 (*Air Pressure*)
'101x003x011',   'Warning',      'Zone 1 CIP - Air pressure is Low',
'101x003x012',   'Warning',      'Zone 2 TriBlender - Air pressure is Low',
'101x003x013',   'Warning',      'Zone 3 Marinade - Air pressure is Low',
'101x003x014',   'Warning',      'Zone 4 Color - Air pressure is Low',

'101x003x021',   'Warning',      'Zone 1 CIP - Air pressure is High',
'101x003x022',   'Warning',      'Zone 2 TriBlender - Air pressure is High',
'101x003x023',   'Warning',      'Zone 3 Marinade - Air pressure is High',
'101x003x024',   'Warning',      'Zone 4 Color - Air pressure is High',

'101x003x111',   'Error',      'Zone 1 CIP - Air pressure is Low',
'101x003x112',   'Error',      'Zone 2 TriBlender - Air pressure is Low',
'101x003x113',   'Error',      'Zone 3 Marinade - Air pressure is Low',
'101x003x114',   'Error',      'Zone 4 Color - Air pressure is Low',

'101x003x121',   'Error',      'Zone 1 CIP - Air pressure is High',
'101x003x122',   'Error',      'Zone 2 TriBlender - Air pressure is High',
'101x003x123',   'Error',      'Zone 3 Marinade - Air pressure is High',
'101x003x124',   'Error',      'Zone 4 Color - Air pressure is High',


  
    (*Emergency*)
'106x001x001',   'Error',      'Emergency cycle 1 (CIP) circuit interrupted',
'106x002x001',   'Error',      'Emergency cycle 2 (Color) circuit interrupted',
'106x003x001',   'Error',      'Emergency cycle 3 (TriBlender) circuit interrupted',
'106x004x001',   'Error',      'Emergency cycle 4 (Marinade) circuit interrupted',

'106x001x002',   'Warning',    'Emergency PB1 Pressed',
'106x002x002',   'Warning',    'Emergency PB2 Pressed',
'106x003x002',   'Warning',    'Emergency PB3_1 Pressed',
'106x003x003',   'Warning',    'Emergency PB3_2 Pressed',
'106x004x002',   'Warning',    'Emergency PB4 Pressed',
'106x000x060',   'Message',    'Emergency Bypass activated',	








    (*Doors*)
	
'107x000x101',   'Warning',    'Door Num 1 Not Closed',
'107x000x102',   'Warning',    'Door Num 2 Not Closed',
'107x000x103',   'Warning',    'Door Num 3 Not Closed',
'107x000x104',   'Warning',    'Door Num 4 Not Closed',

'107x000x121',   'Warning',    'Door Num 1 Not Locked',
'107x000x122',   'Warning',    'Door Num 2 Not Locked',
'107x000x123',   'Warning',    'Door Num 3 Not Locked',
'107x000x124',   'Warning',    'Door Num 4 Not Locked',



    (*Inter lock Zone*)
	
'108x000x141',   'Warning',    'Interlock Zone 1 Robots and Table … doors not locked',
'108x000x142',   'Warning',    'Interlock Zone 2 Load Conveyor … doors not locked',
'108x000x143',   'Warning',    'Interlock Zone 3 Unload Conveyor … doors not locked',
'108x000x144',   'Warning',    'Interlock Zone 4 Manipulator … doors not locked',


      (* Axis ->  FB_Axis *)
'001x000x001',   'Error',   'Motor Power Not OK',
'001x000x002',   'Error',   'Waiting axis reach target',
'001x000x003',   'Error',   'Axis in position check function failed',
'001x000x004',   'Error',   'Limit Detected',
'001x000x005',   'Error',   'Stop Axis',
 

      (* Emergency&Interlock -> prg_Safety *)						  
'002x000x001',   'Error',   'Check EMO devices State',	  
'002x000x002',   'Error',   'TwinSAFE error',	  
'002x000x003',   'Error',   'Check Motors Error',	  
'002x000x004',   'Error',   'check Estop state',	  

 
      (* Initialise -> prg_Initialise *)
'004x000x001',   'Error',   'Wating For Emergency OK',
'004x000x002',   'Error',   'Wating For Interlock OK',
'004x000x003',   'Error',   'Wating For Motors OK',
'004x000x004',   'Error',   'Check Init Station Done',
'004x000x005',   'Error',   'Station Initialization',
'004x000x006',   'Error',   'Loader Initialization',
'004x000x007',   'Error',   'Unload Station',
'004x000x008',   'Error',   'Measuring Station',
'004x000x009',   'Error',   'Gripper Oriantation',
'004x000x010',   'Error',   'index table did not reach home position',
'004x000x012',   'Error',   'carriage position check failed',
'004x000x023',   'Error',   'Wating for Cover Station Init done - check if Robot in safe position',

  

      (* Pneomatic ->  FB_Piston *)
'007x000x001',   'Error',   'Waiting for Sensor Open at Open command',
'007x000x002',   'Error',   'Waiting for Sensor NotClose at Open command',
'007x000x003',   'Error',   'Waiting for Sensor Close at Close command',
'007x000x004',   'Error',   'Waiting for Sensor NotOpen at Close command',
'007x000x005',   'Error',   'No Status',
'007x000x006',   'Error',   'No Valve Operation',
'007x000x007',   'Error',   'Not synchronized with last auto-cycle command',
'007x000x008',   'Error',   'Sensors Checking',

      (* Pneomatic ->  FB_Piston *)
'2AAx001',   'Error',   'Waiting for Sensor Open at Open command',
'2AAx002',   'Error',   'Waiting for Sensor NotClose at Open command',
'2AAx003',   'Error',   'Waiting for Sensor Close at Close command',
'2AAx004',   'Error',   'Waiting for Sensor NotOpen at Close command',
'2AAx005',   'Error',   'No Status',
'2AAx006',   'Error',   'No Valve Operation',
'2AAx007',   'Error',   'Not synchronized with last auto-cycle command',
'2AAx008',   'Error',   'Sensors Checking',	 
		(*Process elementts*)
'109x000x001',   'Warning',   'Conveyor 5 is full',
'109x000x002',   'Error',     'Conveyor 5 is full and Conveyor 4 is ready to output full stack',

'109x000x003',   'Warning',   'Slices Stack is Too Light',
'109x000x004',   'Error',     'Slices Stack is Too Light',

'109x000x005',   'Warning',   'Slices Stack is Too Heavy',
'109x000x006',   'Error',     'Slices Stack is Too Heavy',
 
'555x000x001',   'Error',     'Hello world from NIV',

'985x000x001',   'Warning',     'X lens Constant velocity did not reach during coating',



(*Niv Section*)
(*Cycle X Curtain*)
(*Cycle X & Y*)
(*Cycle X & Theta)
(*Nozzle Operation*)
(*Cycle X Curtain*)
(*Cycle X Curtain*)*)




''];		
END_VAR

// ---- 01 Instance/06-Visu/g_Common.TcGVL
{attribute 'qualified_only'}
VAR_GLOBAL
	iContent_Main: INT;

END_VAR

// ---- 01 Instance/07-Mode/GVL_OperMode.TcGVL
VAR_GLOBAL

	eLightTowerState: E_LightTowerState;
	eBuzzerMode: E_BuzzerMode;
	bBuzzerMute: BOOL;

	bPauseMachine: BOOL;
	bResumeMachine: BOOL;
	bResetAllCycles: BOOL;
	
	PauseAll: BOOL;
	PauseAllDelayed: BOOL;
	ResumeAll: BOOL;	

	iActErrors							: INT;
	iActMessages						: INT;
	iActWarning							: INT;

	fbMode	: ARRAY[0..E_ModeZone.eLast] OF FB_ModeSelect;
	stMode	: ARRAY[0..E_ModeZone.eLast] OF ST_Mode;
	stOper	: ARRAY[0..E_ModeZone.eLast] OF ST_OperationButtons;
	
	fbLightTower: ARRAY[0..E_SkidZone.eLast] OF FB_LightTower;
	fbLightTower_Control: ARRAY[0..E_SkidZone.eLast] OF FB_LightTower_Control;



	//Operational Modes	
	stModeMain: ST_Mode;
	
	// Operational Buttons
	stOpMain				:ST_OperationButtons;
	stOpNonPause			:ST_OperationButtons;	

END_VAR

// ---- 01 Instance/12 Analog Sensor/g_AnalogSensor.TcGVL
//{attribute 'qualified_only'}
VAR_GLOBAL	
	fbAnalogSensor			: ARRAY[0..E_ASense_Name.last] OF FB_AnalogSensor;
	
	//arAnalogSensorName		: ARRAY[0..E_ASense_Name.last] OF STRING(12);
	
	//arAnalogSensorRawValue	: ARRAY[0..E_ASense_Name.last] OF INT;

	iAnalogSensor_sel		: INT:=1;
	
	arAnalogSensorNameList	: ARRAY[0..E_ASense_Name.last] OF STRING(12);
	eAnalogSensorNameList	: E_ASense_Name;

	
END_VAR
//{attribute 'qualified_only'}
VAR_GLOBAL PERSISTENT
	//stAnalogSensorSetting	: ARRAY[0..E_Pis_Name.last] OF ST_Piston_Setting_Param;
	stAnalogSensor			: ARRAY[0..E_ASense_Name.last] OF ST_AnalogSensor;
END_VAR

VAR_GLOBAL CONSTANT

END_VAR

// ---- 01 Instance/13 Process Control/g_ProcControl.TcGVL
//{attribute 'qualified_only'}
VAR_GLOBAL
	//concentration
	(*stDetergent					:	ST_ProcessControl	;
	pcDetergent					: 	FB_ProcessControl	;	//detergent local
	stDisinfectant				:	ST_ProcessControl	;
	pcDisinfectant				: 	FB_ProcessControl	;	//detergent local
    //temperature
	stTemperature_Deterg			:	ST_ProcessControl	;
	pcTemperature_Deterg			: 	FB_ProcessControl	;	//detergent Client	
	stTemperature_Dis				:	ST_ProcessControl	;
	pcTemperature_Dis				: 	FB_ProcessControl	;//disinfectant local/client
	
	//flow rate
	stFlow_Rate						:	ST_ProcessControl	;//CIP
	pcFlow_Rate						: 	FB_ProcessControl	;//disinfectant local/client
	stFlow_Rate_2					:	ST_ProcessControl	;//CLient CIP //level control 
	pcFlow_Rate_2					: 	FB_ProcessControl	;//disinfectant local/client //level control 
	
	//colar marinade 
	//pressure
	stPressure						:	ST_ProcessControl	;
	pcPressure						: 	FB_ProcessControl	;//CIP //Client	
	*)
	
	///////////////////ARRAYS///////////////////
	arr_fbProcCntrl			:	ARRAY [0..E_ProcessControl_Name.eProcCntrl_Last] OF FB_ProcessControl	;
	arr_ProcCntrl_NameList	:	ARRAY [0..E_ProcessControl_Name.eProcCntrl_Last] OF STRING	;
	eProcCntrl_Name			: E_ProcessControl_Name;
END_VAR
VAR_GLOBAL PERSISTENT
	arr_stProcCntrl			:	ARRAY [0..E_ProcessControl_Name.eProcCntrl_Last] OF ST_ProcessControl	;
END_VAR

// ---- 03 Project/30 IO/gIO.TcGVL
//{attribute 'qualified_only'}
VAR_GLOBAL
	i_EL			AT %I*	: ARRAY[1..27] 		OF ST_EL18x9;
	q_EL			AT %Q*	: ARRAY[1..11] 		OF ST_EL28x9;
	ai_EL			AT %I*	: ARRAY[1..6] 		OF ST_EL3xx8;
	aq_EL			AT %Q*	: ARRAY[1..1] 		OF ST_EL4xx8;

	
	q_Manifold1 	AT %Q*	: ARRAY[1..24] 		OF ST_VTUG;
	q_Manifold2 	AT %Q*	: ARRAY[1..24] 		OF ST_VTUG;
	q_Manifold3 	AT %Q*	: ARRAY[1..24] 		OF ST_VTUG;

	Nidec					: ARRAY[0..E_Pump_List.last] 		OF ST_Nidec;

	
	arSafe			: ARRAY[1..1] OF ST_TwinSAFE;
	bStateSafe		: BOOL;
	bStateSafe_ES1	: BOOL;
	bStateSafe_ES2	: BOOL;
	bStateSafe_ES3	: BOOL;
	bStateSafe_ES4	: BOOL;
	
	fbScaleFactor: ARRAY[0..E_ASense_Name.last] 		OF FB_ScaleFactor;
	
	//Anybus Communicator (Box 40), 128 bytes each direction, decoded in g_Anybus.fbAnybus
	Anybus_Inputs_Raw  AT %I* : ARRAY [0..127] OF BYTE;
    Anybus_Outputs_Raw AT %Q* : ARRAY [0..127] OF BYTE;
	Anybus_WcState     AT %I* : BOOL;	//Box 40 WcState, TRUE = process data not valid (also when not in OP)

	
END_VAR

// ---- 03 Project/31 AnybusCommunication/g_Anybus.TcGVL
//{attribute 'qualified_only'}
VAR_GLOBAL
	fbAnybus	: FB_Anybus_Interface;	//CIP <-> Siemens exchange, called in MAIN
	fbSim		: FB_Siemens_Sim;		//Siemens simulator, commissioning only
	bSimEnable	: BOOL;					//TRUE: fbSim replaces the gateway inputs
	arSimRaw	: ARRAY[0..127] OF BYTE;
	bQueueCleared	: BOOL;				//the persistent CIP queue is cleared once after PLC start
	fbBridge	: FB_CIP_Siemens;		//Siemens order -> FB_CIP, CIP state -> Siemens
	bBridgeEnable	: BOOL;				//FALSE: CIP runs from HMI only, stStatus is left alone
END_VAR

// ---- 03 Project/g_Data.TcGVL
//{attribute 'qualified_only'}
VAR_GLOBAL PERSISTENT
	fbCIP						: FB_CIP;
	
	fbCIP_Source				: FB_CIP_Source;
	fbCIP_Return				: FB_CIP_Return;
	fbCIP_Client				: FB_CIP_Client;
	
	arCIP_RequestBufer: ARRAY [0..9] OF ST_CIP_Request;

	//Heat Exchanger
	fbHeatExchenger	:	FB_HeatExchanger	;
	stHeatExchanger	:	ST_HeatExchanger	;
	
	////////////////////////////////////////////////////////////////
	arrTanksSens	:	ARRAY [0..E_Tank_Name.last] OF FB_TankSensors;
	stTanksSens		:	ARRAY [0..E_Tank_Name.last] OF ST_Tank_Level;
	
	////////////////////////////////////////////////////////////////
	arr_CIP_Param		:	ARRAY [0..E_CIP_Usage.eLocal] OF ST_CIP_Param		;//old sets, not read by FB_CIP any more: source of the one-time transfer
	//Recipes of FB_CIP (Vadim 02.11.2026): 0 = Local, 1..30 = CLIENT ID of Siemens
	arr_CIP_Recipe		:	ARRAY [0..cnRecipeMax] OF ST_CIP_Param		;
	arr_CIP_Description	:	ARRAY [0..cnRecipeMax] OF STRING(80)		;//text of the operator, FB_CIP does not read it
	bRecipeTransfer		:	BOOL	;//one-time: old Local, Tank3 Color, Line Color -> recipes 0, 1, 2; reset by MAIN

	//additional variables
	b_CIP_Run	:	BOOL	;
END_VAR
VAR_GLOBAL CONSTANT
	cnRecipeMax			:	INT := 30	;//last recipe = last CLIENT ID
END_VAR

// ---- 00 Library/03 SFC/ITF_FB_SFC_Cycle.TcIO
INTERFACE ITF_FB_SFC_Cycle

METHOD m_Set_SFCFlags_Reference : BOOL
VAR_INPUT
END_VAR
END_METHOD

END_INTERFACE

// ---- 01 Instance/04 Recipe/prg_Call_Recipe_Slow.TcPOU
PROGRAM prg_Call_Recipe_Slow
VAR
	i							: INT;
	bFirstScan					: BOOL:= TRUE;
	ton_RecipeReady				: TON;
	
	
	eRecipeName: E_Recipe_Name;

	r_trigAxisPoints_Loaded: R_TRIG;
	ton_WriteLoaded_Points: TON;
	r_trigRecipe3_loaded: R_TRIG;

	bAllRecipesLoaded: BOOL;
	iRecipeSwitchFrameVar: INT;
	bLoadDefForAll: BOOL;
	
	tPath: STRING(80);
END_VAR

act_Set_StoragePath_For_All();
//act_LoadDeafult();

ton_RecipeReady(PT:=T#1S, IN:=GVL_Recipe.stRecipe[1].bInit AND bFirstScan);
IF ton_RecipeReady.Q THEN;
	bFirstScan:=FALSE;
	bLoadDefForAll:=TRUE;
END_IF




(********************  Other Instances Recipes******************************) // 
FOR eRecipeName:=1 TO E_Recipe_Name.R_Piston_Settings DO	
	fbRecipe[eRecipeName](pstRecipe:=ADR(GVL_Recipe.stRecipe[eRecipeName]), 
			bMemoRecipeUpdated:=, 
			sRecipeDef:=TO_STRING(eRecipeName),
			bLoadDefault:=ar_RecipesLoadDefault[eRecipeName],
			bHMI_FrameActive:=iRecipeSwitchFrameVar=eRecipeName-1,//changed
			sRecipesStoragePath:=ar_RecipesStoragePath[eRecipeName]);
END_FOR
(*			
IF (*fbRecipe_1.bMemoRecipeUpdated AND*) 
fbRecipe_2.bMemoRecipeUpdated 
AND fbRecipe_3.bMemoRecipeUpdated 
AND fbRecipe_4.bMemoRecipeUpdated 
AND fbRecipe_5.bMemoRecipeUpdated 
THEN;
	bAllRecipesLoaded:=TRUE;
ELSE;
	bAllRecipesLoaded:=FALSE;
END_IF
*)

ACTION act_LoadDeafult:
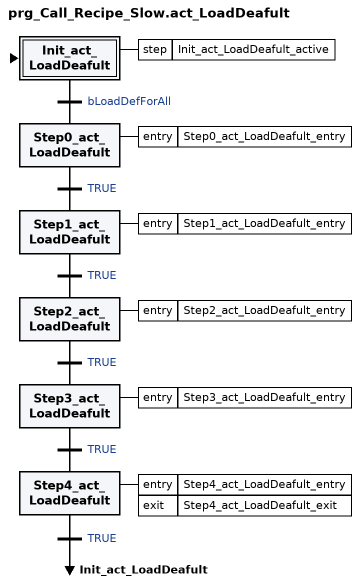
INITIAL_STEP Init_act_LoadDeafult:
    Init_act_LoadDeafult_active(N);  // step action
END_STEP
TRANSITION FROM Init_act_LoadDeafult TO Step0_act_LoadDeafult
    := bLoadDefForAll;
END_TRANSITION
STEP Step0_act_LoadDeafult:  // min time T#2s
    Step0_act_LoadDeafult_entry(P1);  // entry action
END_STEP
TRANSITION FROM Step0_act_LoadDeafult TO Step1_act_LoadDeafult
    := TRUE;
END_TRANSITION
STEP Step1_act_LoadDeafult:  // min time T#2s
    Step1_act_LoadDeafult_entry(P1);  // entry action
END_STEP
TRANSITION FROM Step1_act_LoadDeafult TO Step2_act_LoadDeafult
    := TRUE;
END_TRANSITION
STEP Step2_act_LoadDeafult:  // min time T#2s
    Step2_act_LoadDeafult_entry(P1);  // entry action
END_STEP
TRANSITION FROM Step2_act_LoadDeafult TO Step3_act_LoadDeafult
    := TRUE;
END_TRANSITION
STEP Step3_act_LoadDeafult:  // min time T#2s
    Step3_act_LoadDeafult_entry(P1);  // entry action
END_STEP
TRANSITION FROM Step3_act_LoadDeafult TO Step4_act_LoadDeafult
    := TRUE;
END_TRANSITION
STEP Step4_act_LoadDeafult:  // min time T#2s
    Step4_act_LoadDeafult_entry(P1);  // entry action
    Step4_act_LoadDeafult_exit(P0);  // exit action
END_STEP
TRANSITION FROM Step4_act_LoadDeafult TO Init_act_LoadDeafult
    := TRUE;
END_TRANSITION
END_ACTION

ACTION act_Set_StoragePath_For_All:
FOR eRecipeName:=1 TO E_Recipe_Name.R_Piston_Settings DO;
	GVL_Recipe.ar_RecipesStoragePath_Folder[eRecipeName]:=TO_STRING(eRecipeName);
	tPath:='';
	tPath:=CONCAT(tPath,GVL_Recipe.ar_RecipesStoragePath_Root[GVL_Recipe.eRecipeRootFolder]);
	tPath:=CONCAT(tPath,'\');
	tPath:=CONCAT(tPath,TO_STRING(eRecipeName));
	tPath:=CONCAT(tPath,'\');
	GVL_Recipe.ar_RecipesStoragePath[eRecipeName]:=tPath;
(*
	GVL_Recipe.ar_RecipesStoragePath[eRecipeName]:=
			CONCAT(	GVL_Recipe.ar_RecipesStoragePath_Root[GVL_Recipe.eRecipeRootFolder],'\'); 
	GVL_Recipe.ar_RecipesStoragePath[eRecipeName]:=		
			CONCAT(	GVL_Recipe.ar_RecipesStoragePath[eRecipeName],TO_STRING(eRecipeName));
	GVL_Recipe.ar_RecipesStoragePath[eRecipeName]:=		
			CONCAT(	GVL_Recipe.ar_RecipesStoragePath[eRecipeName],'1');				
	GVL_Recipe.ar_RecipesStoragePath[eRecipeName]:=		
			CONCAT(	GVL_Recipe.ar_RecipesStoragePath[eRecipeName],'\');		
*)	
END_FOR
END_ACTION

ACTION Init_act_LoadDeafult_active:
GVL_Recipe.ar_RecipesLoadDefault[1]:=FALSE;
GVL_Recipe.ar_RecipesLoadDefault[2]:=FALSE;
GVL_Recipe.ar_RecipesLoadDefault[3]:=FALSE;
GVL_Recipe.ar_RecipesLoadDefault[4]:=FALSE;
GVL_Recipe.ar_RecipesLoadDefault[5]:=FALSE;
END_ACTION

ACTION Step0_act_LoadDeafult_entry:
GVL_Recipe.ar_RecipesLoadDefault[1]:=TRUE;
END_ACTION

ACTION Step1_act_LoadDeafult_entry:
GVL_Recipe.ar_RecipesLoadDefault[2]:=TRUE;
END_ACTION

ACTION Step2_act_LoadDeafult_entry:
GVL_Recipe.ar_RecipesLoadDefault[3]:=TRUE;
END_ACTION

ACTION Step3_act_LoadDeafult_entry:
GVL_Recipe.ar_RecipesLoadDefault[4]:=TRUE;
END_ACTION

ACTION Step4_act_LoadDeafult_entry:
GVL_Recipe.ar_RecipesLoadDefault[5]:=TRUE;
END_ACTION

ACTION Step4_act_LoadDeafult_exit:
bLoadDefForAll:=FALSE;
END_ACTION

END_PROGRAM

// ---- POUs/MAIN.TcPOU
PROGRAM MAIN
VAR

	fTotalCIP_Volume: REAL;
	fbWritePersistent: FB_WritePersistentData;
	bTesting		:	BOOL:=FALSE	;
	nI_1			: 	INT		;
	ftg_EStop_Fall	: 	F_TRIG	;
	rs_EStopFall	: 	RS	;
	bTestEstop		:	BOOL:=TRUE	;
	bTemp_Water_Overweight_check: BOOL;
	fbUPS: FB_S_UPS_CX51x0;

END_VAR

prg_RealClock();
prg_Piston();
prg_Safety();
prg_MessageManager();
prg_Messages();
prg_Call_OpMode();
prg_User();
act_ResetPumps();
(*
prg_TriBlender(
		fb_TriBlenderPump:= g_Pump.fbPump[E_Pump_List.TB0001],
		stTriblender:=stTriblender,
		arrComponents:=arrProductionComponents);
*)		
//act_SetAnalogSens_Test();//To be deleted, for testing purposes
act_Call_Sensors_Analog();//To be deleted, for testing purposes
act_Call_Sensors_Analog_1();//To be deleted, for testing purposes
act_Call_ScaleFactor();//To be deleted, for testing purposes
act_Call_ProcessCntrl();

act_Call_Pumps();
act_Sensors();
act_HeatExchenger();
//CIP <-> Siemens exchange
g_Anybus.fbSim(arToCip:=g_Anybus.arSimRaw, arFromCip:=gIO.Anybus_Outputs_Raw);
IF g_Anybus.bSimEnable THEN;
	g_Anybus.fbAnybus(bFieldbusOk:=TRUE, arRawIn:=g_Anybus.arSimRaw, arRawOut:=gIO.Anybus_Outputs_Raw);
ELSE;
	g_Anybus.fbAnybus(bFieldbusOk:=NOT gIO.Anybus_WcState, arRawIn:=gIO.Anybus_Inputs_Raw, arRawOut:=gIO.Anybus_Outputs_Raw);
END_IF
//Requests do not survive a PLC restart (Vadim, 02.11.2026)
IF NOT g_Anybus.bQueueCleared THEN;
	g_Data.fbCIP.m_PosDeleteAll_HMI();
	g_Anybus.bQueueCleared:=TRUE;
END_IF
IF g_Anybus.bBridgeEnable THEN;
	g_Anybus.fbBridge();
	g_Anybus.fbAnybus.stStatus:=g_Anybus.fbBridge.stStatus;
ELSE;
	g_Data.fbCIP.nLocalRecipe:=0;
END_IF
//One-time transfer of the old sets to the new recipes (Vadim 02.11.2026), the rest keeps the program defaults
IF g_Data.bRecipeTransfer THEN;
	g_Data.arr_CIP_Recipe[0]:=g_Data.arr_CIP_Param[E_CIP_Usage.eLocal];
	g_Data.arr_CIP_Recipe[1]:=g_Data.arr_CIP_Param[E_CIP_Usage.eTank_3];
	g_Data.arr_CIP_Recipe[2]:=g_Data.arr_CIP_Param[E_CIP_Usage.eLine_Color];
	g_Data.arr_CIP_Description[0]:='Local';
	g_Data.arr_CIP_Description[1]:='Tank - from Tank3 Color';
	g_Data.arr_CIP_Description[2]:='Pipe - from Line Color';
	g_Data.bRecipeTransfer:=FALSE;
END_IF
act_Call_CIP();

act_Call_For_HMI();

g_SFC.fbSFC_Temp1();

//Temtprary Overweght protection!!!!! DO NOT DELETE
IF fTotalCIP_Volume >=1500 AND FALSE THEN;
	//fbPis[E_Pis_Name.V1022].m_SetByRecipe(stPis:=stPis[E_Pis_Name.V1022], req:=E_Piston_Recipe_State.Release);
	//fbPis[E_Pis_Name.V1019].m_SetByRecipe(stPis:=stPis[E_Pis_Name.V1019], req:=E_Piston_Recipe_State.Release);
	//fbPis[E_Pis_Name.V1016].m_SetByRecipe(stPis:=stPis[E_Pis_Name.V1016], req:=E_Piston_Recipe_State.Release);
	//fbPis[E_Pis_Name.V1011].m_SetByRecipe(stPis:=stPis[E_Pis_Name.V1011], req:=E_Piston_Recipe_State.Release);
	bTemp_Water_Overweight_check:=FALSE;
	fbPrintErrMessageByID(sModuleDescription:='CIP',sActErrorID:='101x000x000');
ELSIF fTotalCIP_Volume < 1480 THEN;
	bTemp_Water_Overweight_check:=TRUE;
END_IF

IF arrTanksSens[E_Tank_Name.T91].get_stTankLevel_OverFlow() THEN;
	fbPis[E_Pis_Name.V1022].m_SetByRecipe(stPis:=stPis[E_Pis_Name.V1022], req:=E_Piston_Recipe_State.Release);
	//print error
	fbPrintErrMessageByID(sModuleDescription:='CIP',sActErrorID:='101x000x001');		
END_IF
IF arrTanksSens[E_Tank_Name.T92].get_stTankLevel_OverFlow() THEN;
	fbPis[E_Pis_Name.V1019].m_SetByRecipe(stPis:=stPis[E_Pis_Name.V1019], req:=E_Piston_Recipe_State.Release);
	//print error
	fbPrintErrMessageByID(sModuleDescription:='CIP',sActErrorID:='101x000x002');		
END_IF
IF arrTanksSens[E_Tank_Name.T93].get_stTankLevel_OverFlow() THEN;
	fbPis[E_Pis_Name.V1016].m_SetByRecipe(stPis:=stPis[E_Pis_Name.V1016], req:=E_Piston_Recipe_State.Release);
	//print error	
	fbPrintErrMessageByID(sModuleDescription:='CIP',sActErrorID:='101x000x003');	
END_IF
IF arrTanksSens[E_Tank_Name.T94].get_stTankLevel_OverFlow() THEN;
	fbPis[E_Pis_Name.V1011].m_SetByRecipe(stPis:=stPis[E_Pis_Name.V1011], req:=E_Piston_Recipe_State.Release);
	//print error
	fbPrintErrMessageByID(sModuleDescription:='CIP',sActErrorID:='101x000x004');		
END_IF
	


mElementList_SetName();

fbWritePersistent(
	NETID:= , 
	PORT:= 851, 
	START:= , 
	TMOUT:= T#3S, 
	MODE:= , 
	BUSY=> , 
	ERR=> , 
	ERRID=> );

fbUPS();

ACTION act_Call_CIP:
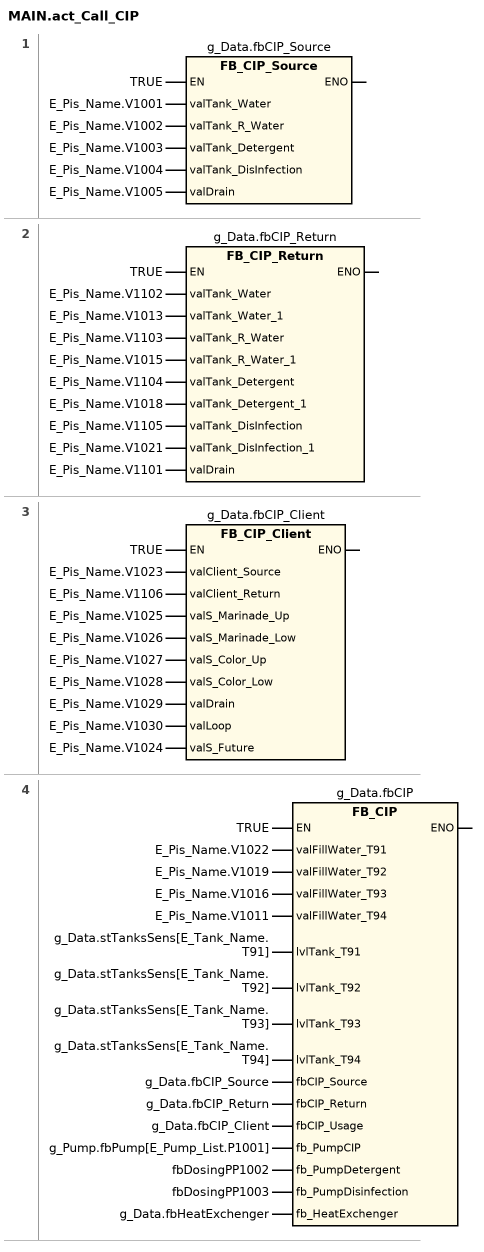
// NETWORK 1
g_Data.fbCIP_Source(
    valTank_Water := E_Pis_Name.V1001,
    valTank_R_Water := E_Pis_Name.V1002,
    valTank_Detergent := E_Pis_Name.V1003,
    valTank_DisInfection := E_Pis_Name.V1004,
    valDrain := E_Pis_Name.V1005); // FB_CIP_Source

// NETWORK 2
g_Data.fbCIP_Return(
    valTank_Water := E_Pis_Name.V1102,
    valTank_Water_1 := E_Pis_Name.V1013,
    valTank_R_Water := E_Pis_Name.V1103,
    valTank_R_Water_1 := E_Pis_Name.V1015,
    valTank_Detergent := E_Pis_Name.V1104,
    valTank_Detergent_1 := E_Pis_Name.V1018,
    valTank_DisInfection := E_Pis_Name.V1105,
    valTank_DisInfection_1 := E_Pis_Name.V1021,
    valDrain := E_Pis_Name.V1101); // FB_CIP_Return

// NETWORK 3
g_Data.fbCIP_Client(
    valClient_Source := E_Pis_Name.V1023,
    valClient_Return := E_Pis_Name.V1106,
    valS_Marinade_Up := E_Pis_Name.V1025,
    valS_Marinade_Low := E_Pis_Name.V1026,
    valS_Color_Up := E_Pis_Name.V1027,
    valS_Color_Low := E_Pis_Name.V1028,
    valDrain := E_Pis_Name.V1029,
    valLoop := E_Pis_Name.V1030,
    valS_Future := E_Pis_Name.V1024); // FB_CIP_Client

// NETWORK 4
g_Data.fbCIP(
    valFillWater_T91 := E_Pis_Name.V1022,
    valFillWater_T92 := E_Pis_Name.V1019,
    valFillWater_T93 := E_Pis_Name.V1016,
    valFillWater_T94 := E_Pis_Name.V1011,
    lvlTank_T91 := g_Data.stTanksSens[E_Tank_Name.T91],
    lvlTank_T92 := g_Data.stTanksSens[E_Tank_Name.T92],
    lvlTank_T93 := g_Data.stTanksSens[E_Tank_Name.T93],
    lvlTank_T94 := g_Data.stTanksSens[E_Tank_Name.T94],
    fbCIP_Source := g_Data.fbCIP_Source,
    fbCIP_Return := g_Data.fbCIP_Return,
    fbCIP_Usage := g_Data.fbCIP_Client,
    fb_PumpCIP := g_Pump.fbPump[E_Pump_List.P1001],
    fb_PumpDetergent := fbDosingPP1002,
    fb_PumpDisinfection := fbDosingPP1003,
    fb_HeatExchenger := g_Data.fbHeatExchenger); // FB_CIP
END_ACTION

ACTION act_Call_For_HMI:


g_HMI.stT91_Sens:=g_Data.stTanksSens[E_Tank_Name.T91];
g_HMI.stT92_Sens:=g_Data.stTanksSens[E_Tank_Name.T92];
g_HMI.stT93_Sens:=g_Data.stTanksSens[E_Tank_Name.T93];
g_HMI.stT94_Sens:=g_Data.stTanksSens[E_Tank_Name.T94];
END_ACTION

ACTION act_Call_ProcessCntrl:
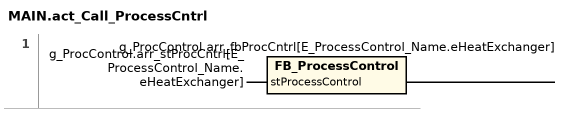
// NETWORK 1
g_ProcControl.arr_fbProcCntrl[E_ProcessControl_Name.eHeatExchanger](stProcessControl := g_ProcControl.arr_stProcCntrl[E_ProcessControl_Name.eHeatExchanger]); // FB_ProcessControl
END_ACTION

ACTION act_Call_Pumps:
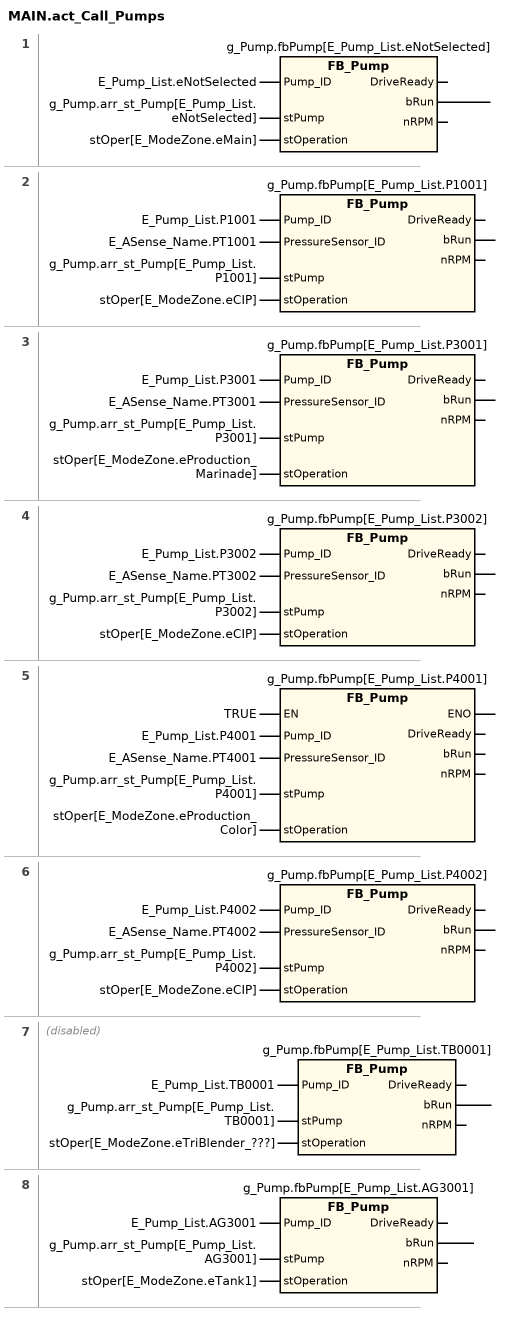
// NETWORK 1
g_Pump.fbPump[E_Pump_List.eNotSelected](
    Pump_ID := E_Pump_List.eNotSelected,
    stPump := g_Pump.arr_st_Pump[E_Pump_List.eNotSelected],
    stOperation := stOper[E_ModeZone.eMain]); // FB_Pump

// NETWORK 2
g_Pump.fbPump[E_Pump_List.P1001](
    Pump_ID := E_Pump_List.P1001,
    PressureSensor_ID := E_ASense_Name.PT1001,
    stPump := g_Pump.arr_st_Pump[E_Pump_List.P1001],
    stOperation := stOper[E_ModeZone.eCIP]); // FB_Pump

// NETWORK 3
g_Pump.fbPump[E_Pump_List.P3001](
    Pump_ID := E_Pump_List.P3001,
    PressureSensor_ID := E_ASense_Name.PT3001,
    stPump := g_Pump.arr_st_Pump[E_Pump_List.P3001],
    stOperation := stOper[E_ModeZone.eProduction_Marinade]); // FB_Pump

// NETWORK 4
g_Pump.fbPump[E_Pump_List.P3002](
    Pump_ID := E_Pump_List.P3002,
    PressureSensor_ID := E_ASense_Name.PT3002,
    stPump := g_Pump.arr_st_Pump[E_Pump_List.P3002],
    stOperation := stOper[E_ModeZone.eCIP]); // FB_Pump

// NETWORK 5
g_Pump.fbPump[E_Pump_List.P4001](
    Pump_ID := E_Pump_List.P4001,
    PressureSensor_ID := E_ASense_Name.PT4001,
    stPump := g_Pump.arr_st_Pump[E_Pump_List.P4001],
    stOperation := stOper[E_ModeZone.eProduction_Color]); // FB_Pump

// NETWORK 6
g_Pump.fbPump[E_Pump_List.P4002](
    Pump_ID := E_Pump_List.P4002,
    PressureSensor_ID := E_ASense_Name.PT4002,
    stPump := g_Pump.arr_st_Pump[E_Pump_List.P4002],
    stOperation := stOper[E_ModeZone.eCIP]); // FB_Pump

// NETWORK 7 (disabled)
// g_Pump.fbPump[E_Pump_List.TB0001](
//     Pump_ID := E_Pump_List.TB0001,
//     stPump := g_Pump.arr_st_Pump[E_Pump_List.TB0001],
//     stOperation := stOper[E_ModeZone.eTriBlender_???]); // FB_Pump

// NETWORK 8
g_Pump.fbPump[E_Pump_List.AG3001](
    Pump_ID := E_Pump_List.AG3001,
    stPump := g_Pump.arr_st_Pump[E_Pump_List.AG3001],
    stOperation := stOper[E_ModeZone.eTank1]); // FB_Pump

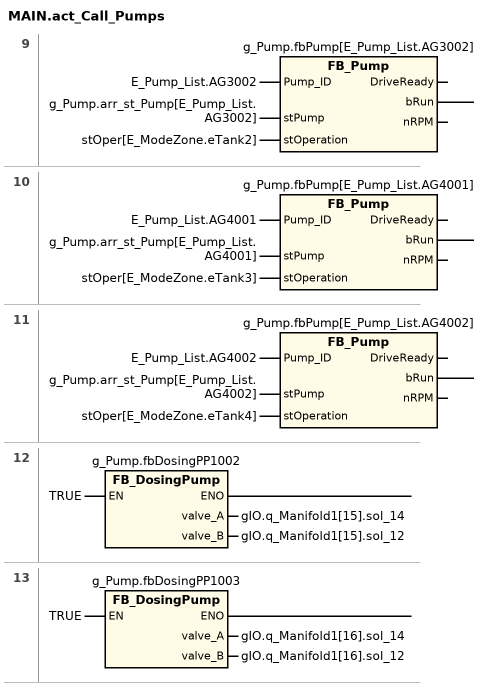
// NETWORK 9
g_Pump.fbPump[E_Pump_List.AG3002](
    Pump_ID := E_Pump_List.AG3002,
    stPump := g_Pump.arr_st_Pump[E_Pump_List.AG3002],
    stOperation := stOper[E_ModeZone.eTank2]); // FB_Pump

// NETWORK 10
g_Pump.fbPump[E_Pump_List.AG4001](
    Pump_ID := E_Pump_List.AG4001,
    stPump := g_Pump.arr_st_Pump[E_Pump_List.AG4001],
    stOperation := stOper[E_ModeZone.eTank3]); // FB_Pump

// NETWORK 11
g_Pump.fbPump[E_Pump_List.AG4002](
    Pump_ID := E_Pump_List.AG4002,
    stPump := g_Pump.arr_st_Pump[E_Pump_List.AG4002],
    stOperation := stOper[E_ModeZone.eTank4]); // FB_Pump

// NETWORK 12
g_Pump.fbDosingPP1002(valve_A => gIO.q_Manifold1[15].sol_14, valve_B => gIO.q_Manifold1[15].sol_12); // FB_DosingPump

// NETWORK 13
g_Pump.fbDosingPP1003(valve_A => gIO.q_Manifold1[16].sol_14, valve_B => gIO.q_Manifold1[16].sol_12); // FB_DosingPump
END_ACTION

ACTION act_Call_ScaleFactor:
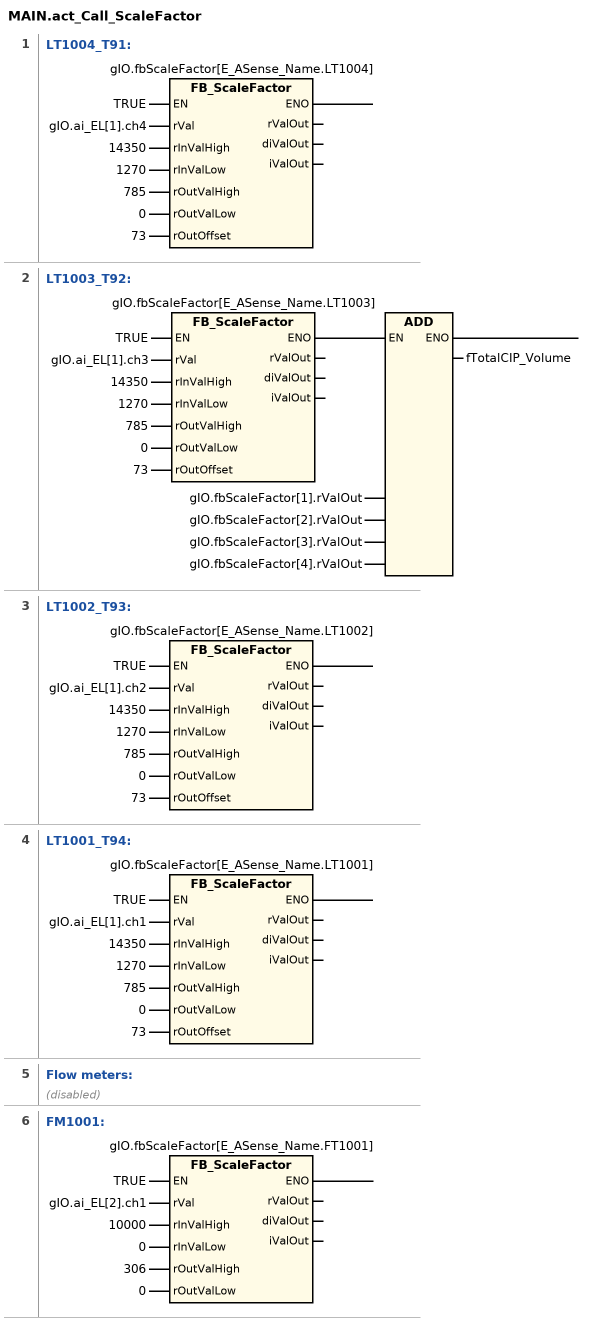
// NETWORK 1
LT1004_T91:
gIO.fbScaleFactor[E_ASense_Name.LT1004](
    rVal := gIO.ai_EL[1].ch4,
    rInValHigh := 14350,
    rInValLow := 1270,
    rOutValHigh := 785,
    rOutValLow := 0,
    rOutOffset := 73); // FB_ScaleFactor

// NETWORK 2
LT1003_T92:
gIO.fbScaleFactor[E_ASense_Name.LT1003](
    rVal := gIO.ai_EL[1].ch3,
    rInValHigh := 14350,
    rInValLow := 1270,
    rOutValHigh := 785,
    rOutValLow := 0,
    rOutOffset := 73); // FB_ScaleFactor
fTotalCIP_Volume := gIO.fbScaleFactor[1].rValOut + gIO.fbScaleFactor[2].rValOut + gIO.fbScaleFactor[3].rValOut + gIO.fbScaleFactor[4].rValOut;

// NETWORK 3
LT1002_T93:
gIO.fbScaleFactor[E_ASense_Name.LT1002](
    rVal := gIO.ai_EL[1].ch2,
    rInValHigh := 14350,
    rInValLow := 1270,
    rOutValHigh := 785,
    rOutValLow := 0,
    rOutOffset := 73); // FB_ScaleFactor

// NETWORK 4
LT1001_T94:
gIO.fbScaleFactor[E_ASense_Name.LT1001](
    rVal := gIO.ai_EL[1].ch1,
    rInValHigh := 14350,
    rInValLow := 1270,
    rOutValHigh := 785,
    rOutValLow := 0,
    rOutOffset := 73); // FB_ScaleFactor

// NETWORK 5 (disabled)
// label: Flow meters

// NETWORK 6
FM1001:
gIO.fbScaleFactor[E_ASense_Name.FT1001](
    rVal := gIO.ai_EL[2].ch1,
    rInValHigh := 10000,
    rInValLow := 0,
    rOutValHigh := 306,
    rOutValLow := 0); // FB_ScaleFactor

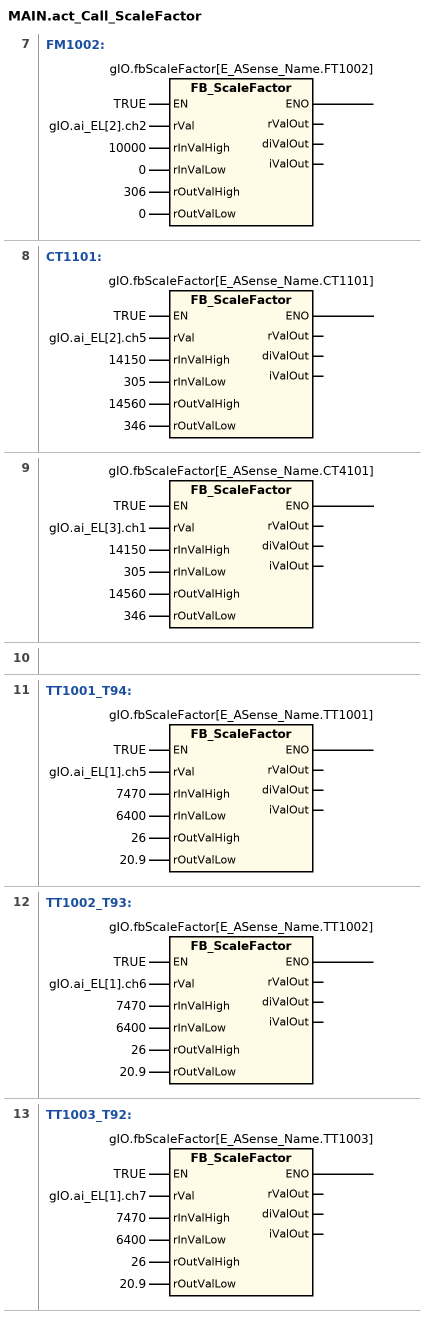
// NETWORK 7
FM1002:
gIO.fbScaleFactor[E_ASense_Name.FT1002](
    rVal := gIO.ai_EL[2].ch2,
    rInValHigh := 10000,
    rInValLow := 0,
    rOutValHigh := 306,
    rOutValLow := 0); // FB_ScaleFactor

// NETWORK 8
CT1101:
gIO.fbScaleFactor[E_ASense_Name.CT1101](
    rVal := gIO.ai_EL[2].ch5,
    rInValHigh := 14150,
    rInValLow := 305,
    rOutValHigh := 14560,
    rOutValLow := 346); // FB_ScaleFactor

// NETWORK 9
gIO.fbScaleFactor[E_ASense_Name.CT4101](
    rVal := gIO.ai_EL[3].ch1,
    rInValHigh := 14150,
    rInValLow := 305,
    rOutValHigh := 14560,
    rOutValLow := 346); // FB_ScaleFactor

// NETWORK 10

// NETWORK 11
TT1001_T94:
gIO.fbScaleFactor[E_ASense_Name.TT1001](
    rVal := gIO.ai_EL[1].ch5,
    rInValHigh := 7470,
    rInValLow := 6400,
    rOutValHigh := 26,
    rOutValLow := 20.9); // FB_ScaleFactor

// NETWORK 12
TT1002_T93:
gIO.fbScaleFactor[E_ASense_Name.TT1002](
    rVal := gIO.ai_EL[1].ch6,
    rInValHigh := 7470,
    rInValLow := 6400,
    rOutValHigh := 26,
    rOutValLow := 20.9); // FB_ScaleFactor

// NETWORK 13
TT1003_T92:
gIO.fbScaleFactor[E_ASense_Name.TT1003](
    rVal := gIO.ai_EL[1].ch7,
    rInValHigh := 7470,
    rInValLow := 6400,
    rOutValHigh := 26,
    rOutValLow := 20.9); // FB_ScaleFactor

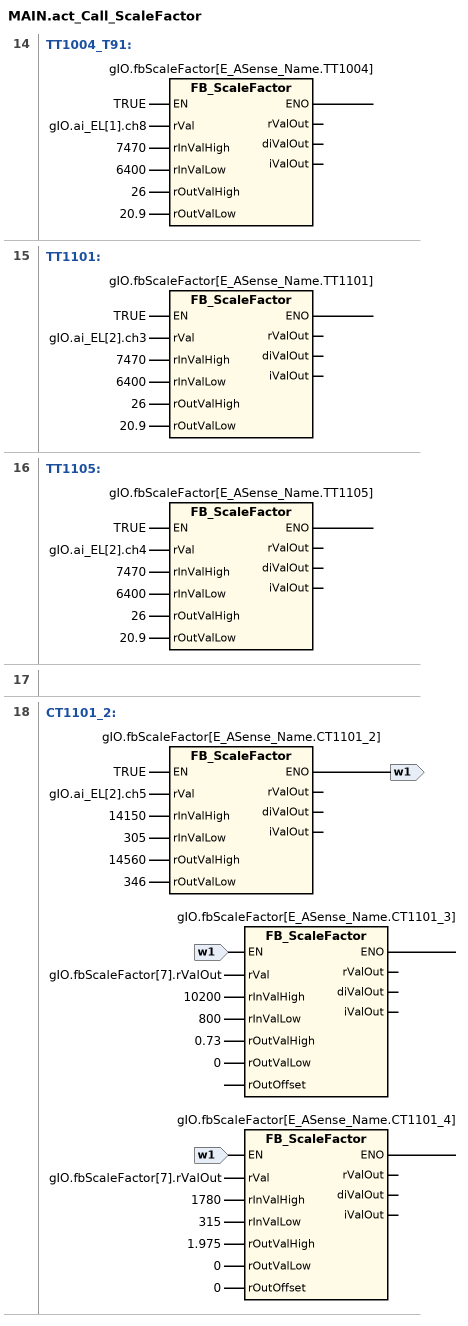
// NETWORK 14
TT1004_T91:
gIO.fbScaleFactor[E_ASense_Name.TT1004](
    rVal := gIO.ai_EL[1].ch8,
    rInValHigh := 7470,
    rInValLow := 6400,
    rOutValHigh := 26,
    rOutValLow := 20.9); // FB_ScaleFactor

// NETWORK 15
TT1101:
gIO.fbScaleFactor[E_ASense_Name.TT1101](
    rVal := gIO.ai_EL[2].ch3,
    rInValHigh := 7470,
    rInValLow := 6400,
    rOutValHigh := 26,
    rOutValLow := 20.9); // FB_ScaleFactor

// NETWORK 16
TT1105:
gIO.fbScaleFactor[E_ASense_Name.TT1105](
    rVal := gIO.ai_EL[2].ch4,
    rInValHigh := 7470,
    rInValLow := 6400,
    rOutValHigh := 26,
    rOutValLow := 20.9); // FB_ScaleFactor

// NETWORK 17

// NETWORK 18
CT1101_2:
gIO.fbScaleFactor[E_ASense_Name.CT1101_2](
    rVal := gIO.ai_EL[2].ch5,
    rInValHigh := 14150,
    rInValLow := 305,
    rOutValHigh := 14560,
    rOutValLow := 346); // FB_ScaleFactor
gIO.fbScaleFactor[E_ASense_Name.CT1101_3](
    rVal := gIO.fbScaleFactor[7].rValOut,
    rInValHigh := 10200,
    rInValLow := 800,
    rOutValHigh := 0.73,
    rOutValLow := 0); // FB_ScaleFactor
gIO.fbScaleFactor[E_ASense_Name.CT1101_4](
    rVal := gIO.fbScaleFactor[7].rValOut,
    rInValHigh := 1780,
    rInValLow := 315,
    rOutValHigh := 1.975,
    rOutValLow := 0,
    rOutOffset := 0); // FB_ScaleFactor

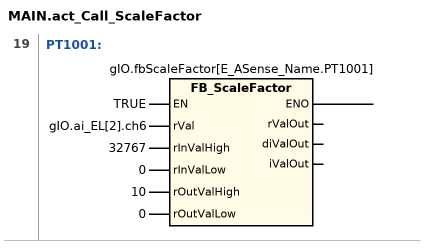
// NETWORK 19
PT1001:
gIO.fbScaleFactor[E_ASense_Name.PT1001](
    rVal := gIO.ai_EL[2].ch6,
    rInValHigh := 32767,
    rInValLow := 0,
    rOutValHigh := 10,
    rOutValLow := 0); // FB_ScaleFactor
END_ACTION

ACTION act_Call_Sensors_Analog:
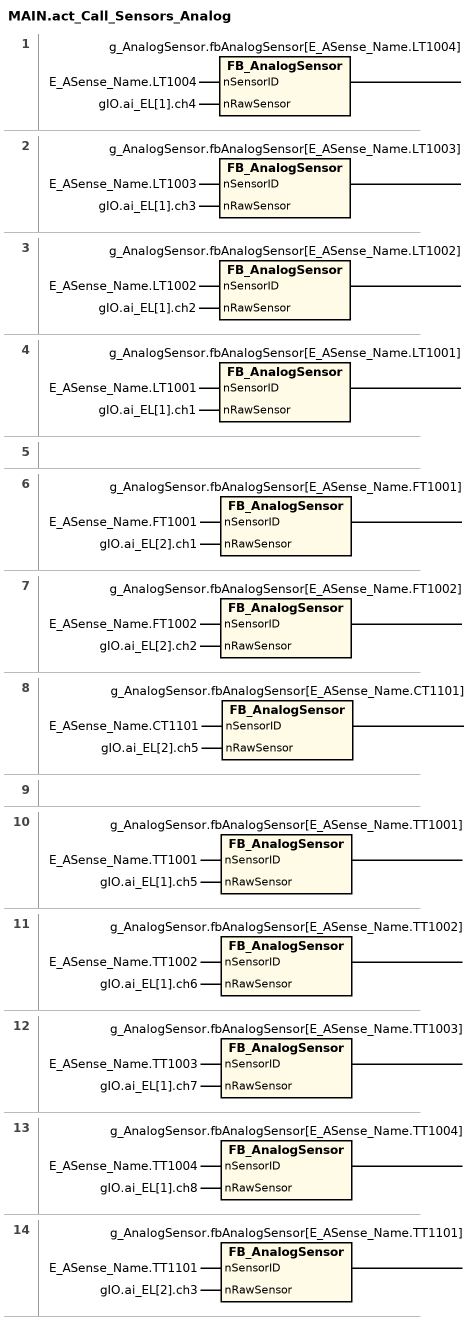
// NETWORK 1
g_AnalogSensor.fbAnalogSensor[E_ASense_Name.LT1004](nSensorID := E_ASense_Name.LT1004, nRawSensor := gIO.ai_EL[1].ch4); // FB_AnalogSensor

// NETWORK 2
g_AnalogSensor.fbAnalogSensor[E_ASense_Name.LT1003](nSensorID := E_ASense_Name.LT1003, nRawSensor := gIO.ai_EL[1].ch3); // FB_AnalogSensor

// NETWORK 3
g_AnalogSensor.fbAnalogSensor[E_ASense_Name.LT1002](nSensorID := E_ASense_Name.LT1002, nRawSensor := gIO.ai_EL[1].ch2); // FB_AnalogSensor

// NETWORK 4
g_AnalogSensor.fbAnalogSensor[E_ASense_Name.LT1001](nSensorID := E_ASense_Name.LT1001, nRawSensor := gIO.ai_EL[1].ch1); // FB_AnalogSensor

// NETWORK 5

// NETWORK 6
g_AnalogSensor.fbAnalogSensor[E_ASense_Name.FT1001](nSensorID := E_ASense_Name.FT1001, nRawSensor := gIO.ai_EL[2].ch1); // FB_AnalogSensor

// NETWORK 7
g_AnalogSensor.fbAnalogSensor[E_ASense_Name.FT1002](nSensorID := E_ASense_Name.FT1002, nRawSensor := gIO.ai_EL[2].ch2); // FB_AnalogSensor

// NETWORK 8
g_AnalogSensor.fbAnalogSensor[E_ASense_Name.CT1101](nSensorID := E_ASense_Name.CT1101, nRawSensor := gIO.ai_EL[2].ch5); // FB_AnalogSensor

// NETWORK 9

// NETWORK 10
g_AnalogSensor.fbAnalogSensor[E_ASense_Name.TT1001](nSensorID := E_ASense_Name.TT1001, nRawSensor := gIO.ai_EL[1].ch5); // FB_AnalogSensor

// NETWORK 11
g_AnalogSensor.fbAnalogSensor[E_ASense_Name.TT1002](nSensorID := E_ASense_Name.TT1002, nRawSensor := gIO.ai_EL[1].ch6); // FB_AnalogSensor

// NETWORK 12
g_AnalogSensor.fbAnalogSensor[E_ASense_Name.TT1003](nSensorID := E_ASense_Name.TT1003, nRawSensor := gIO.ai_EL[1].ch7); // FB_AnalogSensor

// NETWORK 13
g_AnalogSensor.fbAnalogSensor[E_ASense_Name.TT1004](nSensorID := E_ASense_Name.TT1004, nRawSensor := gIO.ai_EL[1].ch8); // FB_AnalogSensor

// NETWORK 14
g_AnalogSensor.fbAnalogSensor[E_ASense_Name.TT1101](nSensorID := E_ASense_Name.TT1101, nRawSensor := gIO.ai_EL[2].ch3); // FB_AnalogSensor

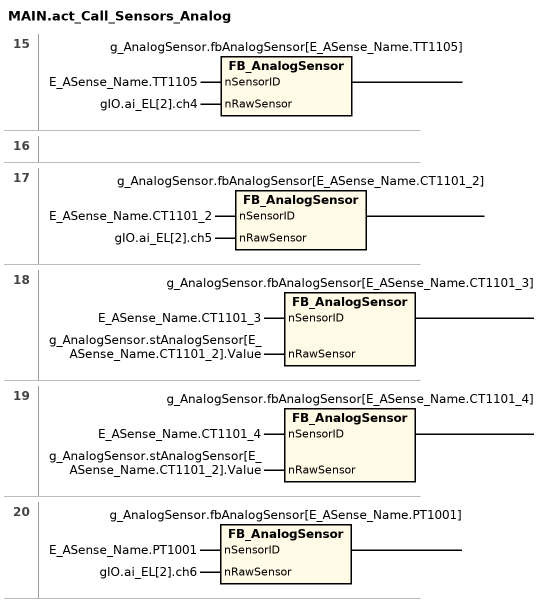
// NETWORK 15
g_AnalogSensor.fbAnalogSensor[E_ASense_Name.TT1105](nSensorID := E_ASense_Name.TT1105, nRawSensor := gIO.ai_EL[2].ch4); // FB_AnalogSensor

// NETWORK 16

// NETWORK 17
g_AnalogSensor.fbAnalogSensor[E_ASense_Name.CT1101_2](nSensorID := E_ASense_Name.CT1101_2, nRawSensor := gIO.ai_EL[2].ch5); // FB_AnalogSensor

// NETWORK 18
g_AnalogSensor.fbAnalogSensor[E_ASense_Name.CT1101_3](nSensorID := E_ASense_Name.CT1101_3, nRawSensor := g_AnalogSensor.stAnalogSensor[E_ASense_Name.CT1101_2].Value); // FB_AnalogSensor

// NETWORK 19
g_AnalogSensor.fbAnalogSensor[E_ASense_Name.CT1101_4](nSensorID := E_ASense_Name.CT1101_4, nRawSensor := g_AnalogSensor.stAnalogSensor[E_ASense_Name.CT1101_2].Value); // FB_AnalogSensor

// NETWORK 20
g_AnalogSensor.fbAnalogSensor[E_ASense_Name.PT1001](nSensorID := E_ASense_Name.PT1001, nRawSensor := gIO.ai_EL[2].ch6); // FB_AnalogSensor
END_ACTION

ACTION act_Call_Sensors_Analog_1:
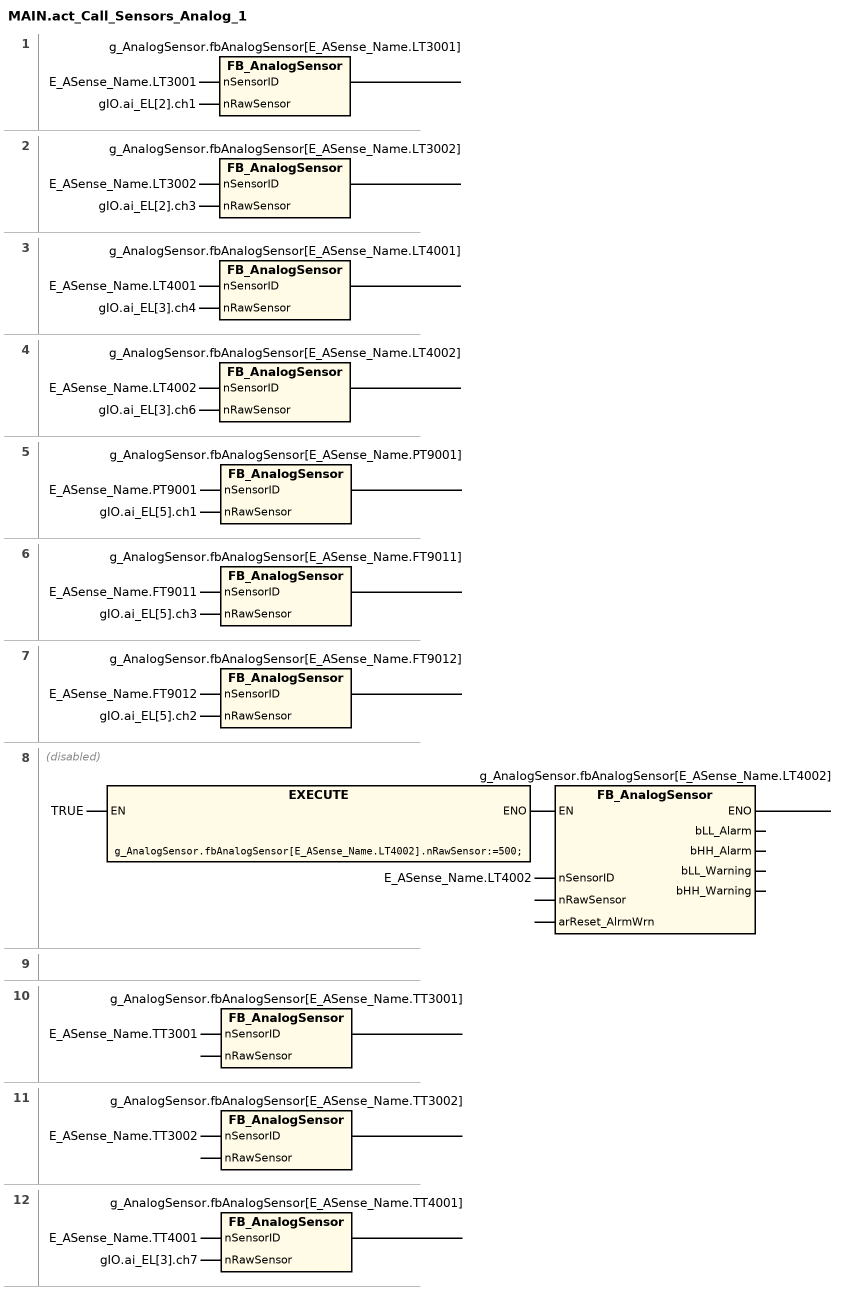
// NETWORK 1
g_AnalogSensor.fbAnalogSensor[E_ASense_Name.LT3001](nSensorID := E_ASense_Name.LT3001, nRawSensor := gIO.ai_EL[2].ch1); // FB_AnalogSensor

// NETWORK 2
g_AnalogSensor.fbAnalogSensor[E_ASense_Name.LT3002](nSensorID := E_ASense_Name.LT3002, nRawSensor := gIO.ai_EL[2].ch3); // FB_AnalogSensor

// NETWORK 3
g_AnalogSensor.fbAnalogSensor[E_ASense_Name.LT4001](nSensorID := E_ASense_Name.LT4001, nRawSensor := gIO.ai_EL[3].ch4); // FB_AnalogSensor

// NETWORK 4
g_AnalogSensor.fbAnalogSensor[E_ASense_Name.LT4002](nSensorID := E_ASense_Name.LT4002, nRawSensor := gIO.ai_EL[3].ch6); // FB_AnalogSensor

// NETWORK 5
g_AnalogSensor.fbAnalogSensor[E_ASense_Name.PT9001](nSensorID := E_ASense_Name.PT9001, nRawSensor := gIO.ai_EL[5].ch1); // FB_AnalogSensor

// NETWORK 6
g_AnalogSensor.fbAnalogSensor[E_ASense_Name.FT9011](nSensorID := E_ASense_Name.FT9011, nRawSensor := gIO.ai_EL[5].ch3); // FB_AnalogSensor

// NETWORK 7
g_AnalogSensor.fbAnalogSensor[E_ASense_Name.FT9012](nSensorID := E_ASense_Name.FT9012, nRawSensor := gIO.ai_EL[5].ch2); // FB_AnalogSensor

// NETWORK 8 (disabled)
// 
// 
// g_AnalogSensor.fbAnalogSensor[E_ASense_Name.LT4002].nRawSensor:=500;
// g_AnalogSensor.fbAnalogSensor[E_ASense_Name.LT4002](nSensorID := E_ASense_Name.LT4002); // FB_AnalogSensor

// NETWORK 9

// NETWORK 10
g_AnalogSensor.fbAnalogSensor[E_ASense_Name.TT3001](nSensorID := E_ASense_Name.TT3001); // FB_AnalogSensor

// NETWORK 11
g_AnalogSensor.fbAnalogSensor[E_ASense_Name.TT3002](nSensorID := E_ASense_Name.TT3002); // FB_AnalogSensor

// NETWORK 12
g_AnalogSensor.fbAnalogSensor[E_ASense_Name.TT4001](nSensorID := E_ASense_Name.TT4001, nRawSensor := gIO.ai_EL[3].ch7); // FB_AnalogSensor

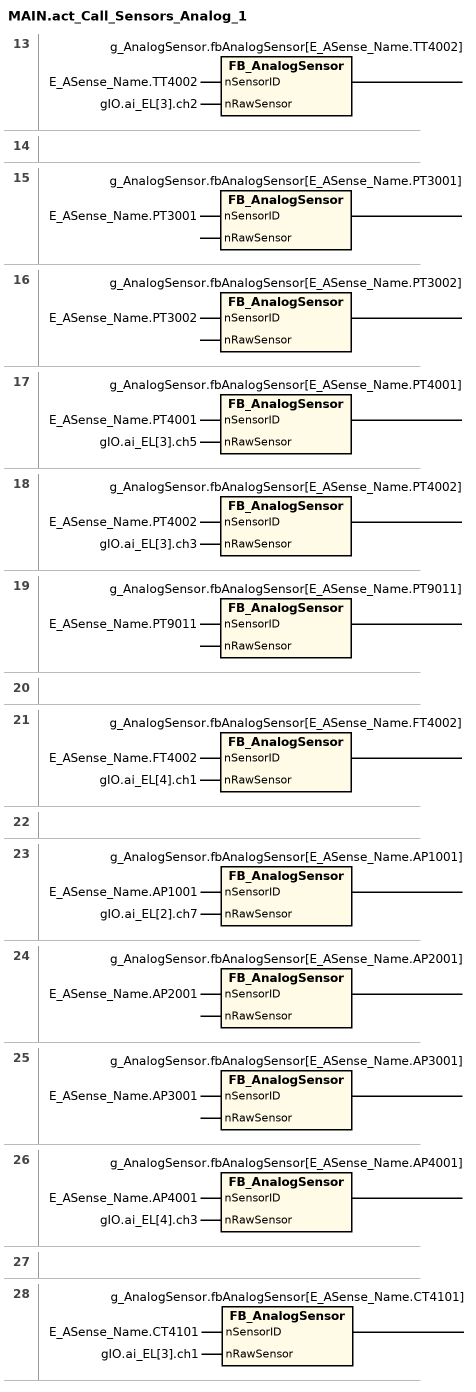
// NETWORK 13
g_AnalogSensor.fbAnalogSensor[E_ASense_Name.TT4002](nSensorID := E_ASense_Name.TT4002, nRawSensor := gIO.ai_EL[3].ch2); // FB_AnalogSensor

// NETWORK 14

// NETWORK 15
g_AnalogSensor.fbAnalogSensor[E_ASense_Name.PT3001](nSensorID := E_ASense_Name.PT3001); // FB_AnalogSensor

// NETWORK 16
g_AnalogSensor.fbAnalogSensor[E_ASense_Name.PT3002](nSensorID := E_ASense_Name.PT3002); // FB_AnalogSensor

// NETWORK 17
g_AnalogSensor.fbAnalogSensor[E_ASense_Name.PT4001](nSensorID := E_ASense_Name.PT4001, nRawSensor := gIO.ai_EL[3].ch5); // FB_AnalogSensor

// NETWORK 18
g_AnalogSensor.fbAnalogSensor[E_ASense_Name.PT4002](nSensorID := E_ASense_Name.PT4002, nRawSensor := gIO.ai_EL[3].ch3); // FB_AnalogSensor

// NETWORK 19
g_AnalogSensor.fbAnalogSensor[E_ASense_Name.PT9011](nSensorID := E_ASense_Name.PT9011); // FB_AnalogSensor

// NETWORK 20

// NETWORK 21
g_AnalogSensor.fbAnalogSensor[E_ASense_Name.FT4002](nSensorID := E_ASense_Name.FT4002, nRawSensor := gIO.ai_EL[4].ch1); // FB_AnalogSensor

// NETWORK 22

// NETWORK 23
g_AnalogSensor.fbAnalogSensor[E_ASense_Name.AP1001](nSensorID := E_ASense_Name.AP1001, nRawSensor := gIO.ai_EL[2].ch7); // FB_AnalogSensor

// NETWORK 24
g_AnalogSensor.fbAnalogSensor[E_ASense_Name.AP2001](nSensorID := E_ASense_Name.AP2001); // FB_AnalogSensor

// NETWORK 25
g_AnalogSensor.fbAnalogSensor[E_ASense_Name.AP3001](nSensorID := E_ASense_Name.AP3001); // FB_AnalogSensor

// NETWORK 26
g_AnalogSensor.fbAnalogSensor[E_ASense_Name.AP4001](nSensorID := E_ASense_Name.AP4001, nRawSensor := gIO.ai_EL[4].ch3); // FB_AnalogSensor

// NETWORK 27

// NETWORK 28
g_AnalogSensor.fbAnalogSensor[E_ASense_Name.CT4101](nSensorID := E_ASense_Name.CT4101, nRawSensor := gIO.ai_EL[3].ch1); // FB_AnalogSensor

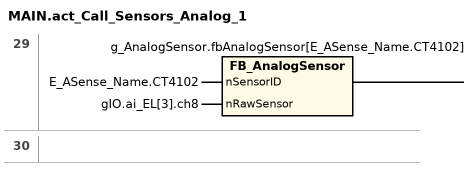
// NETWORK 29
g_AnalogSensor.fbAnalogSensor[E_ASense_Name.CT4102](nSensorID := E_ASense_Name.CT4102, nRawSensor := gIO.ai_EL[3].ch8); // FB_AnalogSensor

// NETWORK 30
END_ACTION

ACTION act_HeatExchenger:
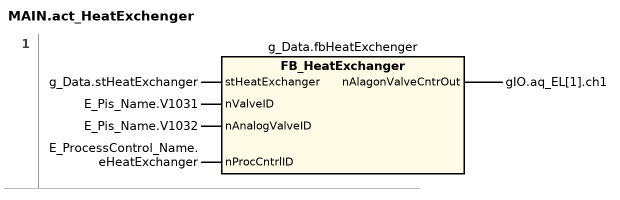
// NETWORK 1
g_Data.fbHeatExchenger(
    stHeatExchanger := g_Data.stHeatExchanger,
    nValveID := E_Pis_Name.V1031,
    nAnalogValveID := E_Pis_Name.V1032,
    nProcCntrlID := E_ProcessControl_Name.eHeatExchanger); // FB_HeatExchanger
gIO.aq_EL[1].ch1 := g_Data.fbHeatExchenger.nAlagonValveCntrOut;
END_ACTION

ACTION act_ResetPumps:
(*ftg_EStop_Fall(CLK:=prg_Safety.ftStateSafe.Q , Q=> );//EStop falling signal
rs_EStopFall(SET:=ftg_EStop_Fall.Q , RESET1:= , Q1=> );
IF rs_EStopFall.Q1 THEN
	FOR nI_1:=1 TO E_Pump_List.last BY 1 DO
		g_Pump.arr_st_Pump[nI_1].bRun_Auto:=FALSE;
	END_FOR
	rs_EStopFall.RESET1:=TRUE;
END_IF
rs_EStopFall.RESET1:=FALSE;*)
;
END_ACTION

ACTION act_Sensors:
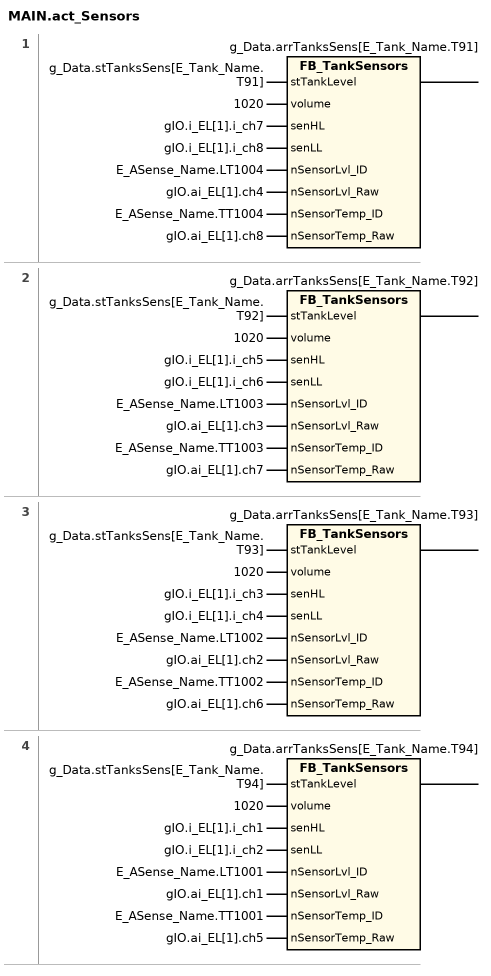
// NETWORK 1
g_Data.arrTanksSens[E_Tank_Name.T91](
    stTankLevel := g_Data.stTanksSens[E_Tank_Name.T91],
    volume := 1020,
    senHL := gIO.i_EL[1].i_ch7,
    senLL := gIO.i_EL[1].i_ch8,
    nSensorLvl_ID := E_ASense_Name.LT1004,
    nSensorLvl_Raw := gIO.ai_EL[1].ch4,
    nSensorTemp_ID := E_ASense_Name.TT1004,
    nSensorTemp_Raw := gIO.ai_EL[1].ch8); // FB_TankSensors

// NETWORK 2
g_Data.arrTanksSens[E_Tank_Name.T92](
    stTankLevel := g_Data.stTanksSens[E_Tank_Name.T92],
    volume := 1020,
    senHL := gIO.i_EL[1].i_ch5,
    senLL := gIO.i_EL[1].i_ch6,
    nSensorLvl_ID := E_ASense_Name.LT1003,
    nSensorLvl_Raw := gIO.ai_EL[1].ch3,
    nSensorTemp_ID := E_ASense_Name.TT1003,
    nSensorTemp_Raw := gIO.ai_EL[1].ch7); // FB_TankSensors

// NETWORK 3
g_Data.arrTanksSens[E_Tank_Name.T93](
    stTankLevel := g_Data.stTanksSens[E_Tank_Name.T93],
    volume := 1020,
    senHL := gIO.i_EL[1].i_ch3,
    senLL := gIO.i_EL[1].i_ch4,
    nSensorLvl_ID := E_ASense_Name.LT1002,
    nSensorLvl_Raw := gIO.ai_EL[1].ch2,
    nSensorTemp_ID := E_ASense_Name.TT1002,
    nSensorTemp_Raw := gIO.ai_EL[1].ch6); // FB_TankSensors

// NETWORK 4
g_Data.arrTanksSens[E_Tank_Name.T94](
    stTankLevel := g_Data.stTanksSens[E_Tank_Name.T94],
    volume := 1020,
    senHL := gIO.i_EL[1].i_ch1,
    senLL := gIO.i_EL[1].i_ch2,
    nSensorLvl_ID := E_ASense_Name.LT1001,
    nSensorLvl_Raw := gIO.ai_EL[1].ch1,
    nSensorTemp_ID := E_ASense_Name.TT1001,
    nSensorTemp_Raw := gIO.ai_EL[1].ch5); // FB_TankSensors
END_ACTION

ACTION act_SetAnalogSens_Test:
//set analog sensors setting only for the test. 
//Later this action should be deleted 
IF NOT bTesting THEN
	//Level
	g_AnalogSensor.stAnalogSensor[E_ASense_Name.LT1004].rawVal_Max:=14350;
	g_AnalogSensor.stAnalogSensor[E_ASense_Name.LT1004].rawVal_Min:=1270;
	g_AnalogSensor.stAnalogSensor[E_ASense_Name.LT1004].outVal_Max:=785;
	g_AnalogSensor.stAnalogSensor[E_ASense_Name.LT1004].outVal_Min:=0;
	g_AnalogSensor.stAnalogSensor[E_ASense_Name.LT1004].outOffset:=73;
	
	g_AnalogSensor.stAnalogSensor[E_ASense_Name.LT1003].rawVal_Max:=14350;
	g_AnalogSensor.stAnalogSensor[E_ASense_Name.LT1003].rawVal_Min:=1270;
	g_AnalogSensor.stAnalogSensor[E_ASense_Name.LT1003].outVal_Max:=785;
	g_AnalogSensor.stAnalogSensor[E_ASense_Name.LT1003].outVal_Min:=0;
	g_AnalogSensor.stAnalogSensor[E_ASense_Name.LT1003].outOffset:=73;
	
	g_AnalogSensor.stAnalogSensor[E_ASense_Name.LT1002].rawVal_Max:=14350;
	g_AnalogSensor.stAnalogSensor[E_ASense_Name.LT1002].rawVal_Min:=1270;
	g_AnalogSensor.stAnalogSensor[E_ASense_Name.LT1002].outVal_Max:=785;
	g_AnalogSensor.stAnalogSensor[E_ASense_Name.LT1002].outVal_Min:=0;
	g_AnalogSensor.stAnalogSensor[E_ASense_Name.LT1002].outOffset:=73;
	
	g_AnalogSensor.stAnalogSensor[E_ASense_Name.LT1001].rawVal_Max:=14350;
	g_AnalogSensor.stAnalogSensor[E_ASense_Name.LT1001].rawVal_Min:=1270;
	g_AnalogSensor.stAnalogSensor[E_ASense_Name.LT1001].outVal_Max:=785;
	g_AnalogSensor.stAnalogSensor[E_ASense_Name.LT1001].outVal_Min:=0;
	g_AnalogSensor.stAnalogSensor[E_ASense_Name.LT1001].outOffset:=73;
	
	//Flow
	g_AnalogSensor.stAnalogSensor[E_ASense_Name.FT1001].rawVal_Max:=10000;
	g_AnalogSensor.stAnalogSensor[E_ASense_Name.FT1001].rawVal_Min:=0;
	g_AnalogSensor.stAnalogSensor[E_ASense_Name.FT1001].outVal_Max:=306;
	g_AnalogSensor.stAnalogSensor[E_ASense_Name.FT1001].outVal_Min:=0;
	g_AnalogSensor.stAnalogSensor[E_ASense_Name.FT1001].outOffset:=0;
	
	g_AnalogSensor.stAnalogSensor[E_ASense_Name.FT1002].rawVal_Max:=10000;
	g_AnalogSensor.stAnalogSensor[E_ASense_Name.FT1002].rawVal_Min:=0;
	g_AnalogSensor.stAnalogSensor[E_ASense_Name.FT1002].outVal_Max:=306;
	g_AnalogSensor.stAnalogSensor[E_ASense_Name.FT1002].outVal_Min:=0;
	g_AnalogSensor.stAnalogSensor[E_ASense_Name.FT1002].outOffset:=0;
	
	////conductivity sensors
	g_AnalogSensor.stAnalogSensor[E_ASense_Name.CT1101].rawVal_Max:=14150;
	g_AnalogSensor.stAnalogSensor[E_ASense_Name.CT1101].rawVal_Min:=305;
	g_AnalogSensor.stAnalogSensor[E_ASense_Name.CT1101].outVal_Max:=14560;
	g_AnalogSensor.stAnalogSensor[E_ASense_Name.CT1101].outVal_Min:=346;
	g_AnalogSensor.stAnalogSensor[E_ASense_Name.CT1101].outOffset:=0;
	(*
	g_AnalogSensor.stAnalogSensor[E_ASense_Name.CT3101].rawVal_Max:=14150;
	g_AnalogSensor.stAnalogSensor[E_ASense_Name.CT3101].rawVal_Min:=305;
	g_AnalogSensor.stAnalogSensor[E_ASense_Name.CT3101].outVal_Max:=14560;
	g_AnalogSensor.stAnalogSensor[E_ASense_Name.CT3101].outVal_Min:=346;
	g_AnalogSensor.stAnalogSensor[E_ASense_Name.CT3101].outOffset:=0;
	*)
	//Temperature sensor
	g_AnalogSensor.stAnalogSensor[E_ASense_Name.TT1001].rawVal_Max:=7470;
	g_AnalogSensor.stAnalogSensor[E_ASense_Name.TT1001].rawVal_Min:=6400;
	g_AnalogSensor.stAnalogSensor[E_ASense_Name.TT1001].outVal_Max:=26;
	g_AnalogSensor.stAnalogSensor[E_ASense_Name.TT1001].outVal_Min:=20.9;
	g_AnalogSensor.stAnalogSensor[E_ASense_Name.TT1001].outOffset:=0;
	
	g_AnalogSensor.stAnalogSensor[E_ASense_Name.TT1002].rawVal_Max:=7470;
	g_AnalogSensor.stAnalogSensor[E_ASense_Name.TT1002].rawVal_Min:=6400;
	g_AnalogSensor.stAnalogSensor[E_ASense_Name.TT1002].outVal_Max:=26;
	g_AnalogSensor.stAnalogSensor[E_ASense_Name.TT1002].outVal_Min:=20.9;
	g_AnalogSensor.stAnalogSensor[E_ASense_Name.TT1002].outOffset:=0;
	
	g_AnalogSensor.stAnalogSensor[E_ASense_Name.TT1003].rawVal_Max:=7470;
	g_AnalogSensor.stAnalogSensor[E_ASense_Name.TT1003].rawVal_Min:=6400;
	g_AnalogSensor.stAnalogSensor[E_ASense_Name.TT1003].outVal_Max:=26;
	g_AnalogSensor.stAnalogSensor[E_ASense_Name.TT1003].outVal_Min:=20.9;
	g_AnalogSensor.stAnalogSensor[E_ASense_Name.TT1003].outOffset:=0;
	
	g_AnalogSensor.stAnalogSensor[E_ASense_Name.TT1004].rawVal_Max:=7470;
	g_AnalogSensor.stAnalogSensor[E_ASense_Name.TT1004].rawVal_Min:=6400;
	g_AnalogSensor.stAnalogSensor[E_ASense_Name.TT1004].outVal_Max:=26;
	g_AnalogSensor.stAnalogSensor[E_ASense_Name.TT1004].outVal_Min:=20.9;
	g_AnalogSensor.stAnalogSensor[E_ASense_Name.TT1004].outOffset:=0;
	
	g_AnalogSensor.stAnalogSensor[E_ASense_Name.TT1101].rawVal_Max:=7470;
	g_AnalogSensor.stAnalogSensor[E_ASense_Name.TT1101].rawVal_Min:=6400;
	g_AnalogSensor.stAnalogSensor[E_ASense_Name.TT1101].outVal_Max:=26;
	g_AnalogSensor.stAnalogSensor[E_ASense_Name.TT1101].outVal_Min:=20.9;
	g_AnalogSensor.stAnalogSensor[E_ASense_Name.TT1101].outOffset:=0;

	bTesting:=TRUE;
END_IF
END_ACTION

METHOD mElementList_SetName : BOOL
VAR_INPUT
END_VAR

VAR
	eASense_Name: E_ASense_Name;
	eProcCntrl: E_ProcessControl_Name;
END_VAR
FOR eASense_Name:=0 TO E_ASense_Name.last DO
	arAnalogSensorNameList[eASense_Name]:=TO_STRING(eASense_Name);
END_FOR

FOR eProcCntrl:=0 TO E_ProcessControl_Name.eProcCntrl_Last DO
	arr_ProcCntrl_NameList[eProcCntrl]:=TO_STRING(eProcCntrl);
	g_ProcControl.arr_stProcCntrl[eProcCntrl].idName:=TO_STRING(eProcCntrl);
END_FOR
END_METHOD

END_PROGRAM

// ---- 00 Library/00-General/TimeAndDate/prg_RealClock.TcPOU
PROGRAM prg_RealClock
VAR

(* Real Time Clock *)
(*	dtRealTime				: DATE_AND_TIME;
	sRealTime				: STRING[22];	
	stSystemTime			: TimeStruct;
	stSystemTime_Empty		: TimeStruct;
	sTime					: STRING[20];
	sDate					: STRING[20];
	sTimeWithMicroSec		: STRING[40];*)

	syncTimer 	: TON;
	fbGetLocalTime 	: NT_GetTime;
	fbRTC_EX2 	: RTC_EX2;
	presetTime 	: TimeStruct;
	syncTrigger 	: F_TRIG;
	bBusy 		: BOOL;
	bError 		: BOOL;
	nErrID 		: UDINT;
	temp1: DATE;
	temp2: TOD;
	NetId :STRING :='';
	bValid_RTCEX2 	: BOOL;
	nMicroseconds 	: DWORD;
	r_trigTrigger: R_TRIG;
	sRealTime_Date	 :STRING(25);
	
	bStartTime: BOOL;
	stStart: TimeStruct;
	sDelta: STRING;
	ton_OneMinuteCount: TON;
END_VAR

(*--------->Set Plc Clock<----------------*)

dtRealTime:=SYSTEMTIME_TO_DT(stSystemTime);
sRealTime:= DT_TO_STRING(dtRealTime);
sRealTime_Date:= DT_TO_STRING(dtRealTime);
sRealTime_Date:=right(sRealTime_Date,19);
temp1:=DT_TO_DATE(dtRealTime);
temp2:=DT_TO_TOD(dtRealTime);
sDate:=DATE_TO_STRING(temp1);
sDate:=DELETE(sDate,2,1);


sTime:=TOD_TO_STRING(temp2);
sTime:=DELETE(sTime,4,1);

sDateTime:=CONCAT(sDate,' ');
sDateTime:=CONCAT(sDateTime,sTime);

sTimeWithMicroSec:=CONCAT(sTime,'.');
sTimeWithMicroSec:=CONCAT(sTimeWithMicroSec,DWORD_TO_STRING(nMicroseconds));




	syncTimer(IN:=NOT SyncTimer.Q , PT:=T#100ms , Q=> , ET=> );
(*r_trigTrigger(CLK:=q_Trigger);*)
	fbGetLocalTime(
		NETID:='' ,
		START:=syncTimer.Q,
		(*START:=r_trigTrigger.Q,*)
		TMOUT:=T#5s ,
		BUSY=>bBusy ,
		ERR=>bError ,
		ERRID=>nErrId ,
		TIMESTR=>presetTime );

	(*syncTrigger(CLK:=NOT bBusy*)
	syncTrigger(CLK:= bBusy
					 AND NOT bError , Q=> );
	fbRTC_EX2(
		EN:=syncTrigger.Q ,
		PDT:=presetTime ,
		PMICRO:=0 ,
		Q=>bValid_RTCEX2 ,
		CDT=>stSystemTime ,
		CMICRO=>nMicroseconds );
		
act_TestDelta();	

ton_OneMinuteCount(PT:=T#1m, IN:=NOT ton_OneMinuteCount.Q);

ACTION act_TestDelta:
IF bStartTime THEN;
	bStartTime:=FALSE;
	stStart:=stSystemTime;
END_IF

sDelta:= m_DeltaTime(stStartTime:=stStart);
END_ACTION

METHOD m_DeltaTime : STRING
VAR_INPUT
	stStartTime  : TimeStruct;
END_VAR
VAR
	tDelta: TIME;
	dtDelta: DATE_AND_TIME;
	todDelta: TOD;


END_VAR
tDelta:=TO_TIME(SYSTEMTIME_TO_DT(stSystemTime)-SYSTEMTIME_TO_DT(stStartTime));

m_DeltaTime:=mTime_to_String_HMI(tInputTime:=tDelta,iSecondDisplay:=FALSE);

(*old
todDelta:=TIME_TO_TOD(tDelta);
m_DeltaTime:=TOD_TO_STRING(todDelta);
m_DeltaTime:=DELETE(m_DeltaTime,4,1);
//dtDelta:=TO_DT(SYSTEMTIME_TO_DT(stSystemTime)-SYSTEMTIME_TO_DT(stStartTime));
//m_DeltaTime:=TIME_TO_STRING(dtDelta);
*)
END_METHOD

METHOD mTime_to_String_HMI : STRING
VAR_INPUT
    tInputTime 		: TIME; // TIME type, stored internally as LTIME (ms)
	iSecondDisplay	: BOOL;
END_VAR
VAR
    nTotalSeconds : UDINT;
    nTotalHours : UDINT;
    nMinutes : UDINT;
    nSeconds : UDINT;
    sFormatted : STRING(20);
END_VAR
// Convert TIME to total seconds
nTotalSeconds := TO_UDINT(tInputTime) / 1000;

// Extract minutes and seconds
nMinutes := nTotalSeconds / 60;
nSeconds := nTotalSeconds MOD 60;

// Convert to total hours
nTotalHours := nMinutes / 60;
nMinutes := nMinutes MOD 60;

// Format output as HHHH:MM:SS (e.g., 0123:45:56)
sFormatted := CONCAT(UDINT_TO_STRING(nTotalHours),'h:');
IF nMinutes < 10 THEN
    sFormatted := CONCAT(sFormatted, '0');
END_IF
sFormatted := CONCAT(sFormatted, UDINT_TO_STRING(nMinutes));
sFormatted := CONCAT(sFormatted, 'm');

IF iSecondDisplay THEN;
	sFormatted := CONCAT(sFormatted, ':');
	IF nSeconds < 10 THEN
		sFormatted := CONCAT(sFormatted, '0');
	END_IF
	sFormatted := CONCAT(sFormatted, UDINT_TO_STRING(nSeconds));
	sFormatted := CONCAT(sFormatted, 's');	
END_IF

// Return formatted string
mTime_to_String_HMI := sFormatted;
END_METHOD

END_PROGRAM

// ---- 01 Instance/01 Piston/prg_Piston.TcPOU
PROGRAM prg_Piston
VAR
	fbPiston: FB_Piston;
	stPiston: ST_Piston;

	bPis_Next_P: BOOL;
	bPis_Next_N: BOOL;

	

	
	TON_0: TON;
	TON_1: TON;
	TON_2: TON;
	TON_3: TON;
	TON_4: TON;
	TON_5: TON;	
	i: INT;
END_VAR

act_InterLock();
act_Call_list_TanksMarinade();
act_Call_list_TanksColor();
act_Call_list_TanksCoolant();
act_Call_List_LineSource();
act_Call_List_LineTarget();
act_Call_list_CIP_SourceNTarget();
act_Call_list_CIP_Client();
act_Call_list_CIP_Tanks();
act_Call_list_Water();
act_Call_list_TriBlender_Selector();


IF bPis_Next_P THEN;
	m_Get_Next_P(iSel:=iPis_sel);
	bPis_Next_P:=FALSE;
END_IF

IF bPis_Next_N THEN;
	m_Get_Next_N(iSel:=iPis_sel);
	bPis_Next_N:=FALSE;
END_IF

FOR i:=0 TO E_Pis_Name.last DO
	ePisNameList:=i;
	arPisNameList[i]:=TO_STRING(ePisNameList);
END_FOR

ACTION act_Call_list_CIP_Client:
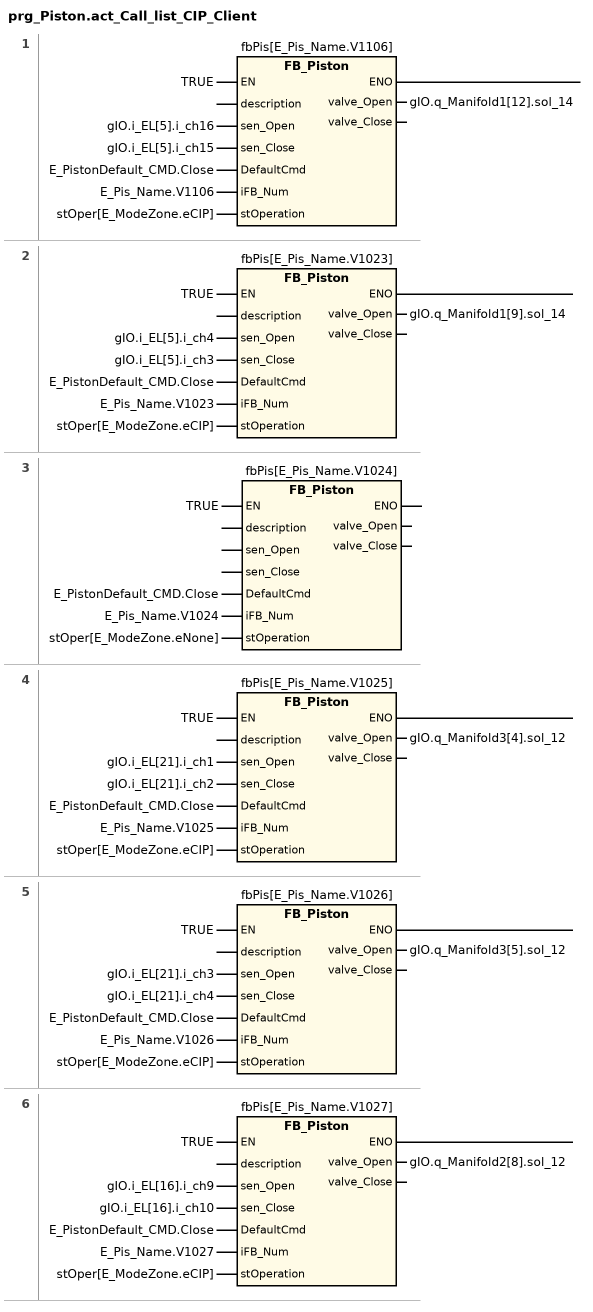
// NETWORK 1
fbPis[E_Pis_Name.V1106](
    sen_Open := gIO.i_EL[5].i_ch16,
    sen_Close := gIO.i_EL[5].i_ch15,
    DefaultCmd := E_PistonDefault_CMD.Close,
    iFB_Num := E_Pis_Name.V1106,
    stOperation := stOper[E_ModeZone.eCIP],
    valve_Open => gIO.q_Manifold1[12].sol_14); // FB_Piston

// NETWORK 2
fbPis[E_Pis_Name.V1023](
    sen_Open := gIO.i_EL[5].i_ch4,
    sen_Close := gIO.i_EL[5].i_ch3,
    DefaultCmd := E_PistonDefault_CMD.Close,
    iFB_Num := E_Pis_Name.V1023,
    stOperation := stOper[E_ModeZone.eCIP],
    valve_Open => gIO.q_Manifold1[9].sol_14); // FB_Piston

// NETWORK 3
fbPis[E_Pis_Name.V1024](
    DefaultCmd := E_PistonDefault_CMD.Close,
    iFB_Num := E_Pis_Name.V1024,
    stOperation := stOper[E_ModeZone.eNone]); // FB_Piston

// NETWORK 4
fbPis[E_Pis_Name.V1025](
    sen_Open := gIO.i_EL[21].i_ch1,
    sen_Close := gIO.i_EL[21].i_ch2,
    DefaultCmd := E_PistonDefault_CMD.Close,
    iFB_Num := E_Pis_Name.V1025,
    stOperation := stOper[E_ModeZone.eCIP],
    valve_Open => gIO.q_Manifold3[4].sol_12); // FB_Piston

// NETWORK 5
fbPis[E_Pis_Name.V1026](
    sen_Open := gIO.i_EL[21].i_ch3,
    sen_Close := gIO.i_EL[21].i_ch4,
    DefaultCmd := E_PistonDefault_CMD.Close,
    iFB_Num := E_Pis_Name.V1026,
    stOperation := stOper[E_ModeZone.eCIP],
    valve_Open => gIO.q_Manifold3[5].sol_12); // FB_Piston

// NETWORK 6
fbPis[E_Pis_Name.V1027](
    sen_Open := gIO.i_EL[16].i_ch9,
    sen_Close := gIO.i_EL[16].i_ch10,
    DefaultCmd := E_PistonDefault_CMD.Close,
    iFB_Num := E_Pis_Name.V1027,
    stOperation := stOper[E_ModeZone.eCIP],
    valve_Open => gIO.q_Manifold2[8].sol_12); // FB_Piston

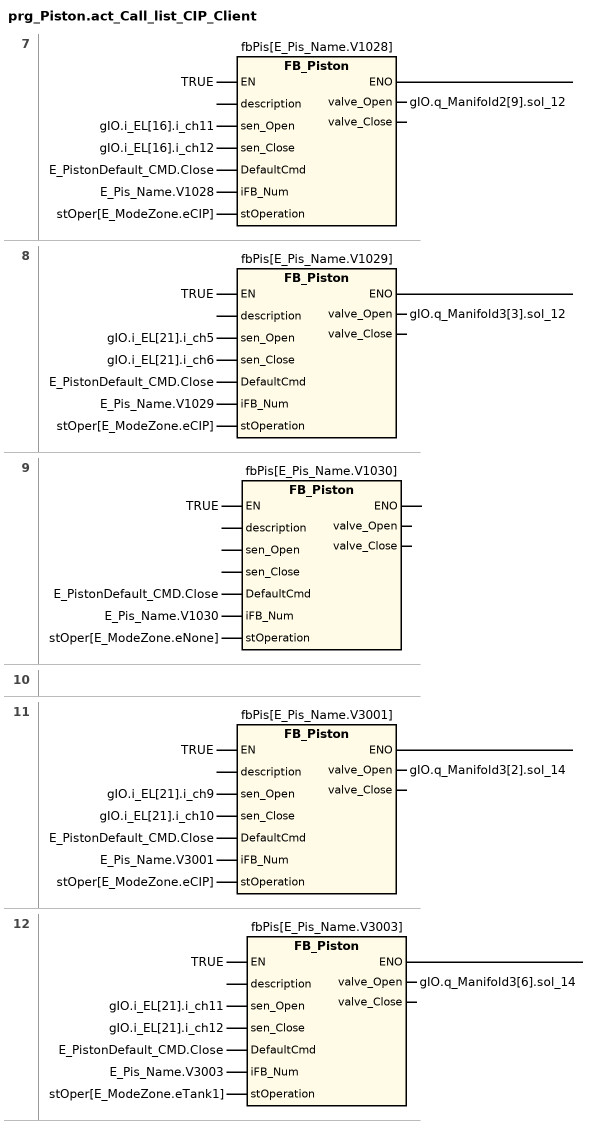
// NETWORK 7
fbPis[E_Pis_Name.V1028](
    sen_Open := gIO.i_EL[16].i_ch11,
    sen_Close := gIO.i_EL[16].i_ch12,
    DefaultCmd := E_PistonDefault_CMD.Close,
    iFB_Num := E_Pis_Name.V1028,
    stOperation := stOper[E_ModeZone.eCIP],
    valve_Open => gIO.q_Manifold2[9].sol_12); // FB_Piston

// NETWORK 8
fbPis[E_Pis_Name.V1029](
    sen_Open := gIO.i_EL[21].i_ch5,
    sen_Close := gIO.i_EL[21].i_ch6,
    DefaultCmd := E_PistonDefault_CMD.Close,
    iFB_Num := E_Pis_Name.V1029,
    stOperation := stOper[E_ModeZone.eCIP],
    valve_Open => gIO.q_Manifold3[3].sol_12); // FB_Piston

// NETWORK 9
fbPis[E_Pis_Name.V1030](
    DefaultCmd := E_PistonDefault_CMD.Close,
    iFB_Num := E_Pis_Name.V1030,
    stOperation := stOper[E_ModeZone.eNone]); // FB_Piston

// NETWORK 10

// NETWORK 11
fbPis[E_Pis_Name.V3001](
    sen_Open := gIO.i_EL[21].i_ch9,
    sen_Close := gIO.i_EL[21].i_ch10,
    DefaultCmd := E_PistonDefault_CMD.Close,
    iFB_Num := E_Pis_Name.V3001,
    stOperation := stOper[E_ModeZone.eCIP],
    valve_Open => gIO.q_Manifold3[2].sol_14); // FB_Piston

// NETWORK 12
fbPis[E_Pis_Name.V3003](
    sen_Open := gIO.i_EL[21].i_ch11,
    sen_Close := gIO.i_EL[21].i_ch12,
    DefaultCmd := E_PistonDefault_CMD.Close,
    iFB_Num := E_Pis_Name.V3003,
    stOperation := stOper[E_ModeZone.eTank1],
    valve_Open => gIO.q_Manifold3[6].sol_14); // FB_Piston

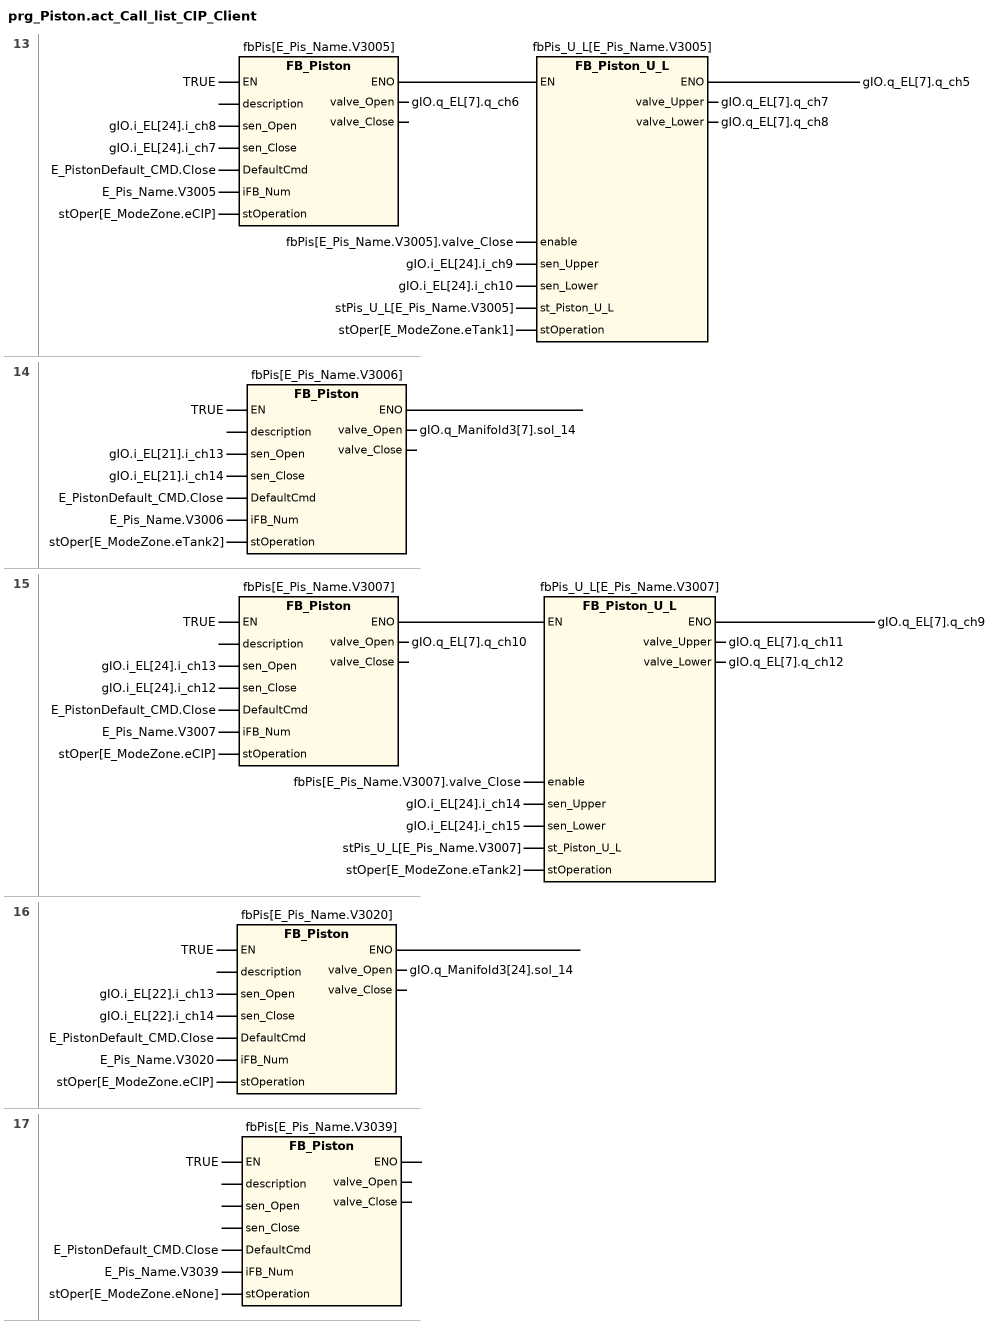
// NETWORK 13
fbPis[E_Pis_Name.V3005](
    sen_Open := gIO.i_EL[24].i_ch8,
    sen_Close := gIO.i_EL[24].i_ch7,
    DefaultCmd := E_PistonDefault_CMD.Close,
    iFB_Num := E_Pis_Name.V3005,
    stOperation := stOper[E_ModeZone.eCIP],
    valve_Open => gIO.q_EL[7].q_ch6); // FB_Piston
fbPis_U_L[E_Pis_Name.V3005](
    enable := fbPis[E_Pis_Name.V3005].valve_Close,
    sen_Upper := gIO.i_EL[24].i_ch9,
    sen_Lower := gIO.i_EL[24].i_ch10,
    st_Piston_U_L := stPis_U_L[E_Pis_Name.V3005],
    stOperation := stOper[E_ModeZone.eTank1],
    valve_Upper => gIO.q_EL[7].q_ch7,
    valve_Lower => gIO.q_EL[7].q_ch8); // FB_Piston_U_L
gIO.q_EL[7].q_ch5 := TRUE;

// NETWORK 14
fbPis[E_Pis_Name.V3006](
    sen_Open := gIO.i_EL[21].i_ch13,
    sen_Close := gIO.i_EL[21].i_ch14,
    DefaultCmd := E_PistonDefault_CMD.Close,
    iFB_Num := E_Pis_Name.V3006,
    stOperation := stOper[E_ModeZone.eTank2],
    valve_Open => gIO.q_Manifold3[7].sol_14); // FB_Piston

// NETWORK 15
fbPis[E_Pis_Name.V3007](
    sen_Open := gIO.i_EL[24].i_ch13,
    sen_Close := gIO.i_EL[24].i_ch12,
    DefaultCmd := E_PistonDefault_CMD.Close,
    iFB_Num := E_Pis_Name.V3007,
    stOperation := stOper[E_ModeZone.eCIP],
    valve_Open => gIO.q_EL[7].q_ch10); // FB_Piston
fbPis_U_L[E_Pis_Name.V3007](
    enable := fbPis[E_Pis_Name.V3007].valve_Close,
    sen_Upper := gIO.i_EL[24].i_ch14,
    sen_Lower := gIO.i_EL[24].i_ch15,
    st_Piston_U_L := stPis_U_L[E_Pis_Name.V3007],
    stOperation := stOper[E_ModeZone.eTank2],
    valve_Upper => gIO.q_EL[7].q_ch11,
    valve_Lower => gIO.q_EL[7].q_ch12); // FB_Piston_U_L
gIO.q_EL[7].q_ch9 := TRUE;

// NETWORK 16
fbPis[E_Pis_Name.V3020](
    sen_Open := gIO.i_EL[22].i_ch13,
    sen_Close := gIO.i_EL[22].i_ch14,
    DefaultCmd := E_PistonDefault_CMD.Close,
    iFB_Num := E_Pis_Name.V3020,
    stOperation := stOper[E_ModeZone.eCIP],
    valve_Open => gIO.q_Manifold3[24].sol_14); // FB_Piston

// NETWORK 17
fbPis[E_Pis_Name.V3039](
    DefaultCmd := E_PistonDefault_CMD.Close,
    iFB_Num := E_Pis_Name.V3039,
    stOperation := stOper[E_ModeZone.eNone]); // FB_Piston

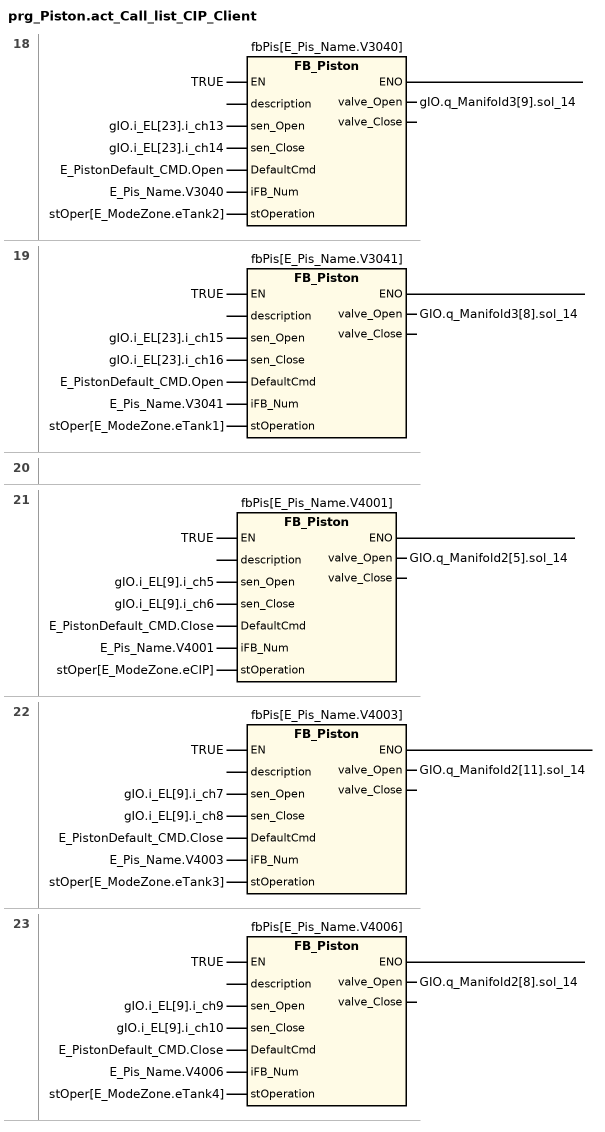
// NETWORK 18
fbPis[E_Pis_Name.V3040](
    sen_Open := gIO.i_EL[23].i_ch13,
    sen_Close := gIO.i_EL[23].i_ch14,
    DefaultCmd := E_PistonDefault_CMD.Open,
    iFB_Num := E_Pis_Name.V3040,
    stOperation := stOper[E_ModeZone.eTank2],
    valve_Open => gIO.q_Manifold3[9].sol_14); // FB_Piston

// NETWORK 19
fbPis[E_Pis_Name.V3041](
    sen_Open := gIO.i_EL[23].i_ch15,
    sen_Close := gIO.i_EL[23].i_ch16,
    DefaultCmd := E_PistonDefault_CMD.Open,
    iFB_Num := E_Pis_Name.V3041,
    stOperation := stOper[E_ModeZone.eTank1],
    valve_Open => GIO.q_Manifold3[8].sol_14); // FB_Piston

// NETWORK 20

// NETWORK 21
fbPis[E_Pis_Name.V4001](
    sen_Open := gIO.i_EL[9].i_ch5,
    sen_Close := gIO.i_EL[9].i_ch6,
    DefaultCmd := E_PistonDefault_CMD.Close,
    iFB_Num := E_Pis_Name.V4001,
    stOperation := stOper[E_ModeZone.eCIP],
    valve_Open => GIO.q_Manifold2[5].sol_14); // FB_Piston

// NETWORK 22
fbPis[E_Pis_Name.V4003](
    sen_Open := gIO.i_EL[9].i_ch7,
    sen_Close := gIO.i_EL[9].i_ch8,
    DefaultCmd := E_PistonDefault_CMD.Close,
    iFB_Num := E_Pis_Name.V4003,
    stOperation := stOper[E_ModeZone.eTank3],
    valve_Open => GIO.q_Manifold2[11].sol_14); // FB_Piston

// NETWORK 23
fbPis[E_Pis_Name.V4006](
    sen_Open := gIO.i_EL[9].i_ch9,
    sen_Close := gIO.i_EL[9].i_ch10,
    DefaultCmd := E_PistonDefault_CMD.Close,
    iFB_Num := E_Pis_Name.V4006,
    stOperation := stOper[E_ModeZone.eTank4],
    valve_Open => GIO.q_Manifold2[8].sol_14); // FB_Piston

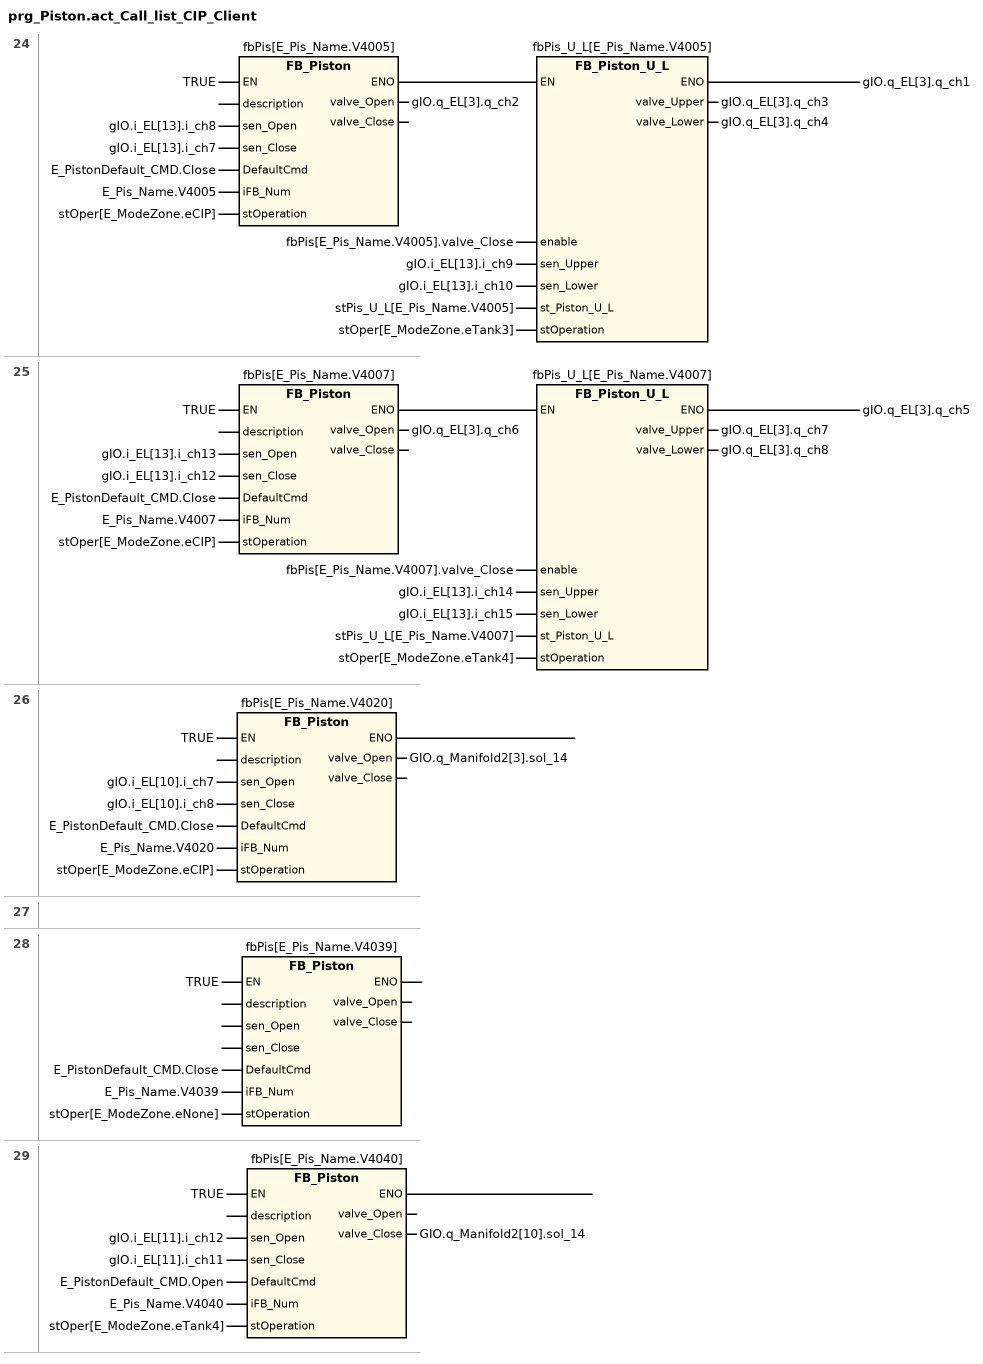
// NETWORK 24
fbPis[E_Pis_Name.V4005](
    sen_Open := gIO.i_EL[13].i_ch8,
    sen_Close := gIO.i_EL[13].i_ch7,
    DefaultCmd := E_PistonDefault_CMD.Close,
    iFB_Num := E_Pis_Name.V4005,
    stOperation := stOper[E_ModeZone.eCIP],
    valve_Open => gIO.q_EL[3].q_ch2); // FB_Piston
fbPis_U_L[E_Pis_Name.V4005](
    enable := fbPis[E_Pis_Name.V4005].valve_Close,
    sen_Upper := gIO.i_EL[13].i_ch9,
    sen_Lower := gIO.i_EL[13].i_ch10,
    st_Piston_U_L := stPis_U_L[E_Pis_Name.V4005],
    stOperation := stOper[E_ModeZone.eTank3],
    valve_Upper => gIO.q_EL[3].q_ch3,
    valve_Lower => gIO.q_EL[3].q_ch4); // FB_Piston_U_L
gIO.q_EL[3].q_ch1 := TRUE;

// NETWORK 25
fbPis[E_Pis_Name.V4007](
    sen_Open := gIO.i_EL[13].i_ch13,
    sen_Close := gIO.i_EL[13].i_ch12,
    DefaultCmd := E_PistonDefault_CMD.Close,
    iFB_Num := E_Pis_Name.V4007,
    stOperation := stOper[E_ModeZone.eCIP],
    valve_Open => gIO.q_EL[3].q_ch6); // FB_Piston
fbPis_U_L[E_Pis_Name.V4007](
    enable := fbPis[E_Pis_Name.V4007].valve_Close,
    sen_Upper := gIO.i_EL[13].i_ch14,
    sen_Lower := gIO.i_EL[13].i_ch15,
    st_Piston_U_L := stPis_U_L[E_Pis_Name.V4007],
    stOperation := stOper[E_ModeZone.eTank4],
    valve_Upper => gIO.q_EL[3].q_ch7,
    valve_Lower => gIO.q_EL[3].q_ch8); // FB_Piston_U_L
gIO.q_EL[3].q_ch5 := TRUE;

// NETWORK 26
fbPis[E_Pis_Name.V4020](
    sen_Open := gIO.i_EL[10].i_ch7,
    sen_Close := gIO.i_EL[10].i_ch8,
    DefaultCmd := E_PistonDefault_CMD.Close,
    iFB_Num := E_Pis_Name.V4020,
    stOperation := stOper[E_ModeZone.eCIP],
    valve_Open => GIO.q_Manifold2[3].sol_14); // FB_Piston

// NETWORK 27

// NETWORK 28
fbPis[E_Pis_Name.V4039](
    DefaultCmd := E_PistonDefault_CMD.Close,
    iFB_Num := E_Pis_Name.V4039,
    stOperation := stOper[E_ModeZone.eNone]); // FB_Piston

// NETWORK 29
fbPis[E_Pis_Name.V4040](
    sen_Open := gIO.i_EL[11].i_ch12,
    sen_Close := gIO.i_EL[11].i_ch11,
    DefaultCmd := E_PistonDefault_CMD.Open,
    iFB_Num := E_Pis_Name.V4040,
    stOperation := stOper[E_ModeZone.eTank4],
    valve_Close => GIO.q_Manifold2[10].sol_14); // FB_Piston

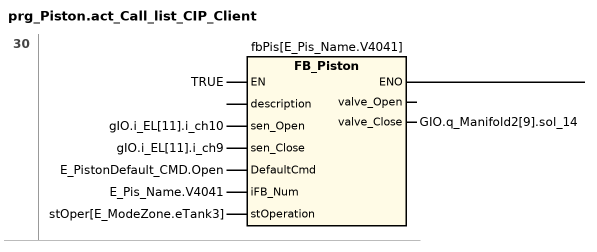
// NETWORK 30
fbPis[E_Pis_Name.V4041](
    sen_Open := gIO.i_EL[11].i_ch10,
    sen_Close := gIO.i_EL[11].i_ch9,
    DefaultCmd := E_PistonDefault_CMD.Open,
    iFB_Num := E_Pis_Name.V4041,
    stOperation := stOper[E_ModeZone.eTank3],
    valve_Close => GIO.q_Manifold2[9].sol_14); // FB_Piston
END_ACTION

ACTION act_Call_list_CIP_SourceNTarget:
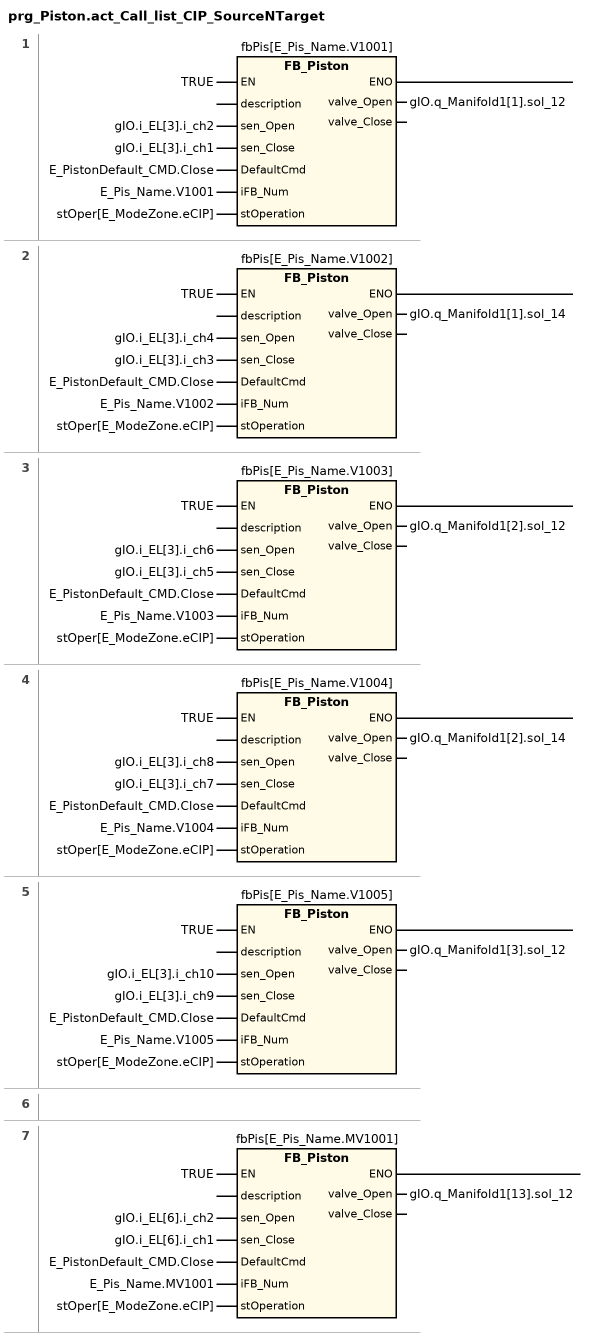
// NETWORK 1
fbPis[E_Pis_Name.V1001](
    sen_Open := gIO.i_EL[3].i_ch2,
    sen_Close := gIO.i_EL[3].i_ch1,
    DefaultCmd := E_PistonDefault_CMD.Close,
    iFB_Num := E_Pis_Name.V1001,
    stOperation := stOper[E_ModeZone.eCIP],
    valve_Open => gIO.q_Manifold1[1].sol_12); // FB_Piston

// NETWORK 2
fbPis[E_Pis_Name.V1002](
    sen_Open := gIO.i_EL[3].i_ch4,
    sen_Close := gIO.i_EL[3].i_ch3,
    DefaultCmd := E_PistonDefault_CMD.Close,
    iFB_Num := E_Pis_Name.V1002,
    stOperation := stOper[E_ModeZone.eCIP],
    valve_Open => gIO.q_Manifold1[1].sol_14); // FB_Piston

// NETWORK 3
fbPis[E_Pis_Name.V1003](
    sen_Open := gIO.i_EL[3].i_ch6,
    sen_Close := gIO.i_EL[3].i_ch5,
    DefaultCmd := E_PistonDefault_CMD.Close,
    iFB_Num := E_Pis_Name.V1003,
    stOperation := stOper[E_ModeZone.eCIP],
    valve_Open => gIO.q_Manifold1[2].sol_12); // FB_Piston

// NETWORK 4
fbPis[E_Pis_Name.V1004](
    sen_Open := gIO.i_EL[3].i_ch8,
    sen_Close := gIO.i_EL[3].i_ch7,
    DefaultCmd := E_PistonDefault_CMD.Close,
    iFB_Num := E_Pis_Name.V1004,
    stOperation := stOper[E_ModeZone.eCIP],
    valve_Open => gIO.q_Manifold1[2].sol_14); // FB_Piston

// NETWORK 5
fbPis[E_Pis_Name.V1005](
    sen_Open := gIO.i_EL[3].i_ch10,
    sen_Close := gIO.i_EL[3].i_ch9,
    DefaultCmd := E_PistonDefault_CMD.Close,
    iFB_Num := E_Pis_Name.V1005,
    stOperation := stOper[E_ModeZone.eCIP],
    valve_Open => gIO.q_Manifold1[3].sol_12); // FB_Piston

// NETWORK 6

// NETWORK 7
fbPis[E_Pis_Name.MV1001](
    sen_Open := gIO.i_EL[6].i_ch2,
    sen_Close := gIO.i_EL[6].i_ch1,
    DefaultCmd := E_PistonDefault_CMD.Close,
    iFB_Num := E_Pis_Name.MV1001,
    stOperation := stOper[E_ModeZone.eCIP],
    valve_Open => gIO.q_Manifold1[13].sol_12); // FB_Piston

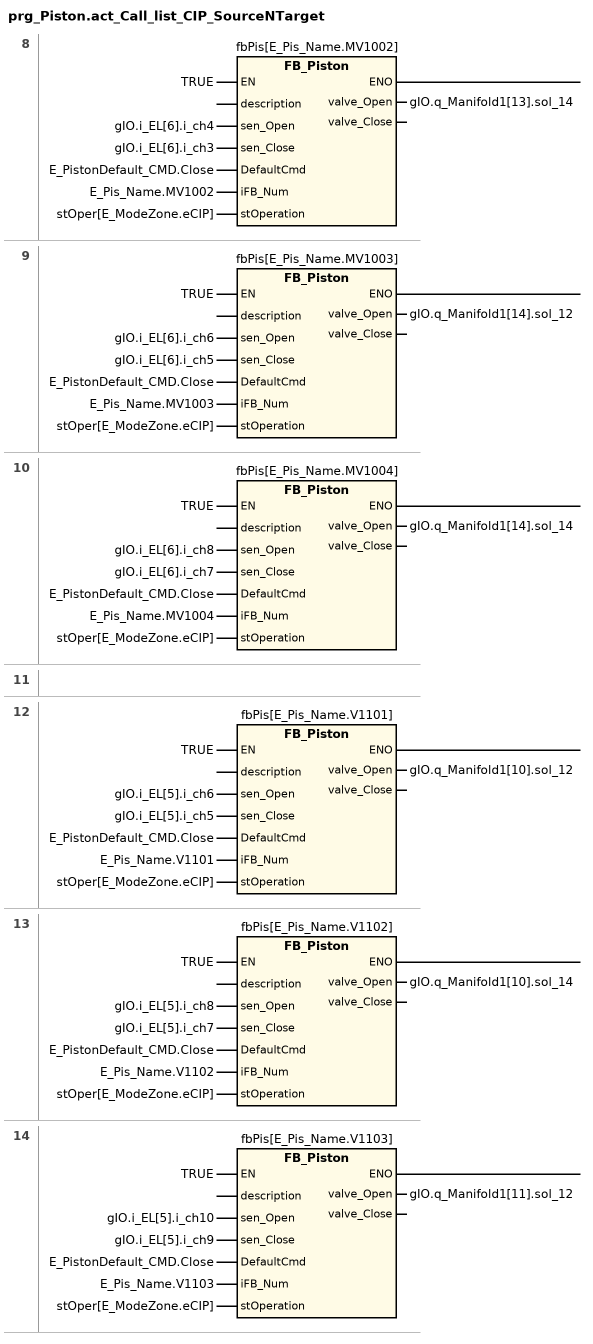
// NETWORK 8
fbPis[E_Pis_Name.MV1002](
    sen_Open := gIO.i_EL[6].i_ch4,
    sen_Close := gIO.i_EL[6].i_ch3,
    DefaultCmd := E_PistonDefault_CMD.Close,
    iFB_Num := E_Pis_Name.MV1002,
    stOperation := stOper[E_ModeZone.eCIP],
    valve_Open => gIO.q_Manifold1[13].sol_14); // FB_Piston

// NETWORK 9
fbPis[E_Pis_Name.MV1003](
    sen_Open := gIO.i_EL[6].i_ch6,
    sen_Close := gIO.i_EL[6].i_ch5,
    DefaultCmd := E_PistonDefault_CMD.Close,
    iFB_Num := E_Pis_Name.MV1003,
    stOperation := stOper[E_ModeZone.eCIP],
    valve_Open => gIO.q_Manifold1[14].sol_12); // FB_Piston

// NETWORK 10
fbPis[E_Pis_Name.MV1004](
    sen_Open := gIO.i_EL[6].i_ch8,
    sen_Close := gIO.i_EL[6].i_ch7,
    DefaultCmd := E_PistonDefault_CMD.Close,
    iFB_Num := E_Pis_Name.MV1004,
    stOperation := stOper[E_ModeZone.eCIP],
    valve_Open => gIO.q_Manifold1[14].sol_14); // FB_Piston

// NETWORK 11

// NETWORK 12
fbPis[E_Pis_Name.V1101](
    sen_Open := gIO.i_EL[5].i_ch6,
    sen_Close := gIO.i_EL[5].i_ch5,
    DefaultCmd := E_PistonDefault_CMD.Close,
    iFB_Num := E_Pis_Name.V1101,
    stOperation := stOper[E_ModeZone.eCIP],
    valve_Open => gIO.q_Manifold1[10].sol_12); // FB_Piston

// NETWORK 13
fbPis[E_Pis_Name.V1102](
    sen_Open := gIO.i_EL[5].i_ch8,
    sen_Close := gIO.i_EL[5].i_ch7,
    DefaultCmd := E_PistonDefault_CMD.Close,
    iFB_Num := E_Pis_Name.V1102,
    stOperation := stOper[E_ModeZone.eCIP],
    valve_Open => gIO.q_Manifold1[10].sol_14); // FB_Piston

// NETWORK 14
fbPis[E_Pis_Name.V1103](
    sen_Open := gIO.i_EL[5].i_ch10,
    sen_Close := gIO.i_EL[5].i_ch9,
    DefaultCmd := E_PistonDefault_CMD.Close,
    iFB_Num := E_Pis_Name.V1103,
    stOperation := stOper[E_ModeZone.eCIP],
    valve_Open => gIO.q_Manifold1[11].sol_12); // FB_Piston

